REGION Network 21: Transition for STATE Num:60 StWtL1S2DownOver
   RUNG wire#powerrail
      Contact( #sStWtL1S2DownOver )
      I_Contact( #sStWtResetRel )
      Contact( #sSst )
      Contact( #iL1S2DownOver )
      Coil( #sStWtL1S2DownOver_T1 )
   END_RUNG
   // the same network as SCL:
   #sStWtL1S2DownOver_T1 := #sStWtL1S2DownOver AND NOT #sStWtResetRel AND #sSst AND #iL1S2DownOver;
END_REGION

REGION Network 22: STATE Num:60 StWtL1S2DownOver
   RUNG wire#powerrail
      Contact( #sStWtL1S2DownOver )
      wire#w1
      I_Contact( #sStWtResetRel )
      I_Contact( #sStWtL1S2DownOver_T1 )
      wire#w2
      Coil( #sStWtL1S2DownOver )
   END_RUNG
   RUNG wire#powerrail
      Contact( #sStWtLifterAtPos1_T1 )
   END_RUNG wire#w1
   RUNG wire#powerrail
      Contact( #sStRecovery_T7 )
   END_RUNG wire#w1
   RUNG wire#w2
      { S7_GenerateENO := "TRUE" } Move(in := 60, out1 => #StateNo)
   END_RUNG
   // the same network as SCL:
   #sStWtL1S2DownOver := (#sStWtL1S2DownOver OR #sStWtLifterAtPos1_T1 OR #sStRecovery_T7) AND NOT #sStWtResetRel AND NOT #sStWtL1S2DownOver_T1;
   IF #sStWtL1S2DownOver THEN #StateNo := 60; END_IF;
END_REGION

REGION Network 23: Actions for STATE Num:60 StWtL1S2DownOver
   RUNG wire#powerrail
      Contact( #sStWtL1S2DownOver )
      Coil( #qL1S2Down )
   END_RUNG
   // the same network as SCL:
   #qL1S2Down := #sStWtL1S2DownOver;
END_REGION

REGION Network 24: Transition for STATE Num:70 StWtOTSFrmConv
   RUNG wire#powerrail
      Contact( #sStWtOTSFrmConv )
      I_Contact( #sStWtResetRel )
      Contact( #sSst )
      Contact( #iOTSFrmConv )
      Coil( #sStWtOTSFrmConv_T1 )
   END_RUNG
   // the same network as SCL:
   #sStWtOTSFrmConv_T1 := #sStWtOTSFrmConv AND NOT #sStWtResetRel AND #sSst AND #iOTSFrmConv;
END_REGION

REGION Network 25: STATE Num:70 StWtOTSFrmConv
   RUNG wire#powerrail
      Contact( #sStWtOTSFrmConv )
      wire#w1
      I_Contact( #sStWtResetRel )
      I_Contact( #sStWtOTSFrmConv_T1 )
      wire#w2
      Coil( #sStWtOTSFrmConv )
   END_RUNG
   RUNG wire#powerrail
      Contact( #sStWtL1S2DownOver_T1 )
   END_RUNG wire#w1
   RUNG wire#w2
      { S7_GenerateENO := "TRUE" } Move(in := 70, out1 => #StateNo)
   END_RUNG
   // the same network as SCL:
   #sStWtOTSFrmConv := (#sStWtOTSFrmConv OR #sStWtL1S2DownOver_T1) AND NOT #sStWtResetRel AND NOT #sStWtOTSFrmConv_T1;
   IF #sStWtOTSFrmConv THEN #StateNo := 70; END_IF;
END_REGION

REGION Network 26: Actions for STATE Num:70 StWtOTSFrmConv
   RUNG wire#powerrail
      Contact( #sStWtOTSFrmConv )
      Coil( #qRTRToConv )
   END_RUNG
   // the same network as SCL:
   #qRTRToConv := #sStWtOTSFrmConv;
END_REGION

REGION Network 27: Transition for STATE Num:80 StWtL1RecvBegin
   RUNG wire#powerrail
      Contact( #sStWtL1RecvBegin )
      I_Contact( #sStWtResetRel )
      Contact( #sSst )
      I_Contact( #iReceiveAreaClear )
      Coil( #sStWtL1RecvBegin_T1 )
   END_RUNG
   // the same network as SCL:
   #sStWtL1RecvBegin_T1 := #sStWtL1RecvBegin AND NOT #sStWtResetRel AND #sSst AND NOT #iReceiveAreaClear;
END_REGION

REGION Network 28: STATE Num:80 StWtL1RecvBegin
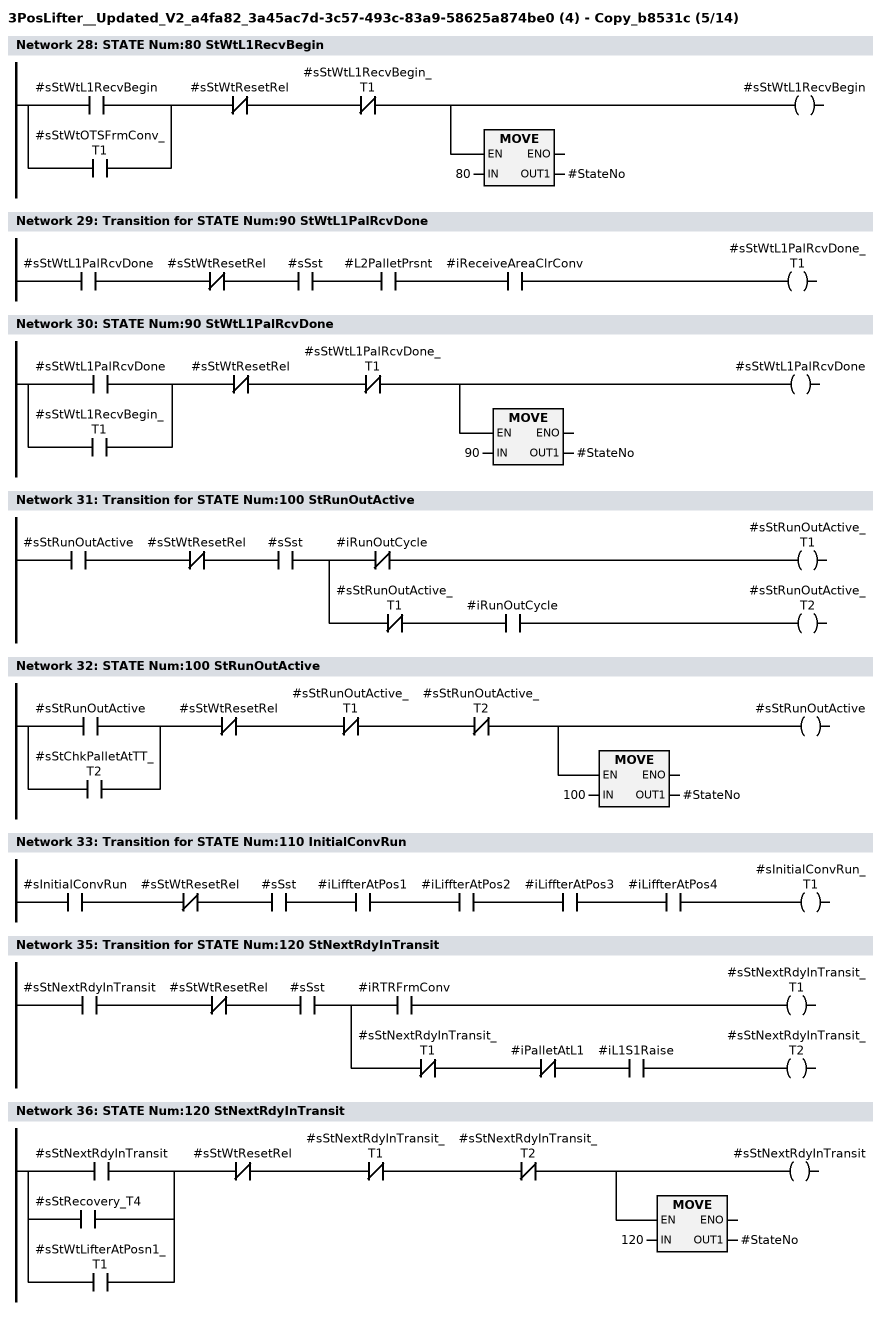
   RUNG wire#powerrail
      Contact( #sStWtL1RecvBegin )
      wire#w1
      I_Contact( #sStWtResetRel )
      I_Contact( #sStWtL1RecvBegin_T1 )
      wire#w2
      Coil( #sStWtL1RecvBegin )
   END_RUNG
   RUNG wire#powerrail
      Contact( #sStWtOTSFrmConv_T1 )
   END_RUNG wire#w1
   RUNG wire#w2
      { S7_GenerateENO := "TRUE" } Move(in := 80, out1 => #StateNo)
   END_RUNG
   // the same network as SCL:
   #sStWtL1RecvBegin := (#sStWtL1RecvBegin OR #sStWtOTSFrmConv_T1) AND NOT #sStWtResetRel AND NOT #sStWtL1RecvBegin_T1;
   IF #sStWtL1RecvBegin THEN #StateNo := 80; END_IF;
END_REGION

REGION Network 29: Transition for STATE Num:90 StWtL1PalRcvDone
   RUNG wire#powerrail
      Contact( #sStWtL1PalRcvDone )
      I_Contact( #sStWtResetRel )
      Contact( #sSst )
      Contact( #L2PalletPrsnt )
      Contact( #iReceiveAreaClrConv )
      Coil( #sStWtL1PalRcvDone_T1 )
   END_RUNG
   // the same network as SCL:
   #sStWtL1PalRcvDone_T1 := #sStWtL1PalRcvDone AND NOT #sStWtResetRel AND #sSst AND #L2PalletPrsnt AND #iReceiveAreaClrConv;
END_REGION

REGION Network 30: STATE Num:90 StWtL1PalRcvDone
   RUNG wire#powerrail
      Contact( #sStWtL1PalRcvDone )
      wire#w1
      I_Contact( #sStWtResetRel )
      I_Contact( #sStWtL1PalRcvDone_T1 )
      wire#w2
      Coil( #sStWtL1PalRcvDone )
   END_RUNG
   RUNG wire#powerrail
      Contact( #sStWtL1RecvBegin_T1 )
   END_RUNG wire#w1
   RUNG wire#w2
      { S7_GenerateENO := "TRUE" } Move(in := 90, out1 => #StateNo)
   END_RUNG
   // the same network as SCL:
   #sStWtL1PalRcvDone := (#sStWtL1PalRcvDone OR #sStWtL1RecvBegin_T1) AND NOT #sStWtResetRel AND NOT #sStWtL1PalRcvDone_T1;
   IF #sStWtL1PalRcvDone THEN #StateNo := 90; END_IF;
END_REGION

REGION Network 31: Transition for STATE Num:100 StRunOutActive
   RUNG wire#powerrail
      Contact( #sStRunOutActive )
      I_Contact( #sStWtResetRel )
      Contact( #sSst )
      wire#w1
      I_Contact( #iRunOutCycle )
      Coil( #sStRunOutActive_T1 )
   END_RUNG
   RUNG wire#w1
      I_Contact( #sStRunOutActive_T1 )
      Contact( #iRunOutCycle )
      Coil( #sStRunOutActive_T2 )
   END_RUNG
   // the same network as SCL:
   #_w1 := #sStRunOutActive AND NOT #sStWtResetRel AND #sSst;
   #sStRunOutActive_T1 := #_w1 AND NOT #iRunOutCycle;
   #sStRunOutActive_T2 := #_w1 AND NOT #sStRunOutActive_T1 AND #iRunOutCycle;
END_REGION

REGION Network 32: STATE Num:100 StRunOutActive
   RUNG wire#powerrail
      Contact( #sStRunOutActive )
      wire#w1
      I_Contact( #sStWtResetRel )
      I_Contact( #sStRunOutActive_T1 )
      I_Contact( #sStRunOutActive_T2 )
      wire#w2
      Coil( #sStRunOutActive )
   END_RUNG
   RUNG wire#powerrail
      Contact( #sStChkPalletAtTT_T2 )
   END_RUNG wire#w1
   RUNG wire#w2
      { S7_GenerateENO := "TRUE" } Move(in := 100, out1 => #StateNo)
   END_RUNG
   // the same network as SCL:
   #sStRunOutActive := (#sStRunOutActive OR #sStChkPalletAtTT_T2) AND NOT #sStWtResetRel AND NOT #sStRunOutActive_T1 AND NOT #sStRunOutActive_T2;
   IF #sStRunOutActive THEN #StateNo := 100; END_IF;
END_REGION

REGION Network 33: Transition for STATE Num:110 InitialConvRun
   RUNG wire#powerrail
      Contact( #sInitialConvRun )
      I_Contact( #sStWtResetRel )
      Contact( #sSst )
      Contact( #iLiffterAtPos1 )
      Contact( #iLiffterAtPos2 )
      Contact( #iLiffterAtPos3 )
      Contact( #iLiffterAtPos4 )
      Coil( #sInitialConvRun_T1 )
   END_RUNG
   // the same network as SCL:
   #sInitialConvRun_T1 := #sInitialConvRun AND NOT #sStWtResetRel AND #sSst AND #iLiffterAtPos1 AND #iLiffterAtPos2 AND #iLiffterAtPos3 AND #iLiffterAtPos4;
END_REGION

NETWORK
TITLE = STATE Num:110 InitialConvRun
      A(;
      O     #sInitialConvRun;
//wrong transition variable removed
      );
      AN    #sStWtResetRel;
      AN    #sInitialConvRun_T1;
      =     %L1.0;
      A     %L1.0;
      BLD   102;
      =     #sInitialConvRun;
      A     %L1.0;
      JNB   Label_110;
      L     110;
      T     #StateNo;
Label_110:NOP   0;

REGION Network 35: Transition for STATE Num:120 StNextRdyInTransit
   RUNG wire#powerrail
      Contact( #sStNextRdyInTransit )
      I_Contact( #sStWtResetRel )
      Contact( #sSst )
      wire#w1
      Contact( #iRTRFrmConv )
      Coil( #sStNextRdyInTransit_T1 )
   END_RUNG
   RUNG wire#w1
      I_Contact( #sStNextRdyInTransit_T1 )
      I_Contact( #iPalletAtL1 )
      Contact( #iL1S1Raise )
      Coil( #sStNextRdyInTransit_T2 )
   END_RUNG
   // the same network as SCL:
   #_w1 := #sStNextRdyInTransit AND NOT #sStWtResetRel AND #sSst;
   #sStNextRdyInTransit_T1 := #_w1 AND #iRTRFrmConv;
   #sStNextRdyInTransit_T2 := #_w1 AND NOT #sStNextRdyInTransit_T1 AND NOT #iPalletAtL1 AND #iL1S1Raise;
END_REGION

REGION Network 36: STATE Num:120 StNextRdyInTransit
   RUNG wire#powerrail
      Contact( #sStNextRdyInTransit )
      wire#w1
      I_Contact( #sStWtResetRel )
      I_Contact( #sStNextRdyInTransit_T1 )
      I_Contact( #sStNextRdyInTransit_T2 )
      wire#w2
      Coil( #sStNextRdyInTransit )
   END_RUNG
   RUNG wire#powerrail
      Contact( #sStRecovery_T4 )
   END_RUNG wire#w1
   RUNG wire#powerrail
      Contact( #sStWtLifterAtPosn1_T1 )
   END_RUNG wire#w1
   RUNG wire#w2
      { S7_GenerateENO := "TRUE" } Move(in := 120, out1 => #StateNo)
   END_RUNG
   // the same network as SCL:
   #sStNextRdyInTransit := (#sStNextRdyInTransit OR #sStRecovery_T4 OR #sStWtLifterAtPosn1_T1) AND NOT #sStWtResetRel AND NOT #sStNextRdyInTransit_T1 AND NOT #sStNextRdyInTransit_T2;
   IF #sStNextRdyInTransit THEN #StateNo := 120; END_IF;
END_REGION

REGION Network 37: Transition for STATE Num:130 StNextRdyInTransit_1
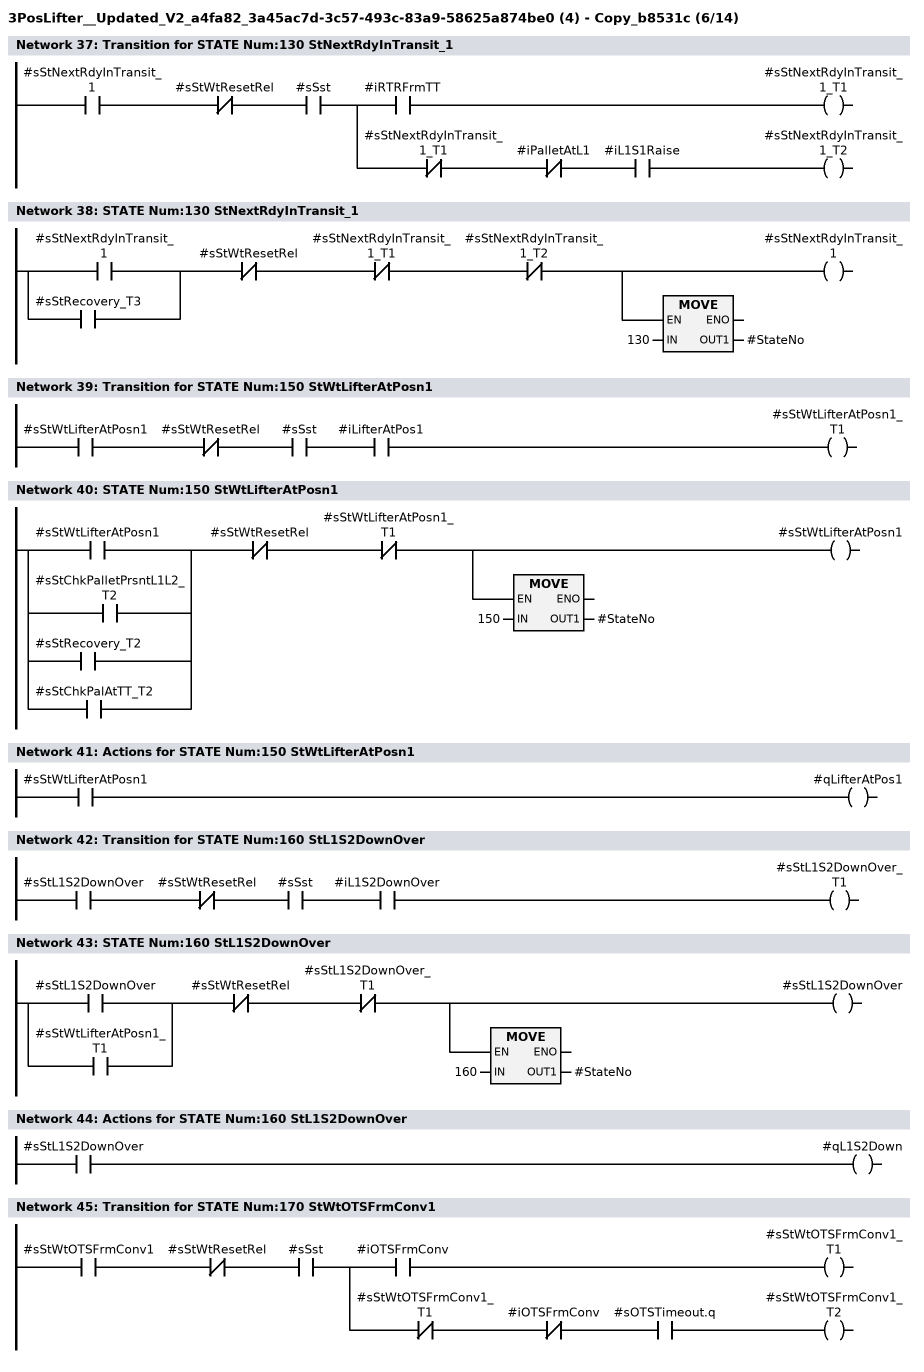
   RUNG wire#powerrail
      Contact( #sStNextRdyInTransit_1 )
      I_Contact( #sStWtResetRel )
      Contact( #sSst )
      wire#w1
      Contact( #iRTRFrmTT )
      Coil( #sStNextRdyInTransit_1_T1 )
   END_RUNG
   RUNG wire#w1
      I_Contact( #sStNextRdyInTransit_1_T1 )
      I_Contact( #iPalletAtL1 )
      Contact( #iL1S1Raise )
      Coil( #sStNextRdyInTransit_1_T2 )
   END_RUNG
   // the same network as SCL:
   #_w1 := #sStNextRdyInTransit_1 AND NOT #sStWtResetRel AND #sSst;
   #sStNextRdyInTransit_1_T1 := #_w1 AND #iRTRFrmTT;
   #sStNextRdyInTransit_1_T2 := #_w1 AND NOT #sStNextRdyInTransit_1_T1 AND NOT #iPalletAtL1 AND #iL1S1Raise;
END_REGION

REGION Network 38: STATE Num:130 StNextRdyInTransit_1
   RUNG wire#powerrail
      Contact( #sStNextRdyInTransit_1 )
      wire#w1
      I_Contact( #sStWtResetRel )
      I_Contact( #sStNextRdyInTransit_1_T1 )
      I_Contact( #sStNextRdyInTransit_1_T2 )
      wire#w2
      Coil( #sStNextRdyInTransit_1 )
   END_RUNG
   RUNG wire#powerrail
      Contact( #sStRecovery_T3 )
   END_RUNG wire#w1
   RUNG wire#w2
      { S7_GenerateENO := "TRUE" } Move(in := 130, out1 => #StateNo)
   END_RUNG
   // the same network as SCL:
   #sStNextRdyInTransit_1 := (#sStNextRdyInTransit_1 OR #sStRecovery_T3) AND NOT #sStWtResetRel AND NOT #sStNextRdyInTransit_1_T1 AND NOT #sStNextRdyInTransit_1_T2;
   IF #sStNextRdyInTransit_1 THEN #StateNo := 130; END_IF;
END_REGION

REGION Network 39: Transition for STATE Num:150 StWtLifterAtPosn1
   RUNG wire#powerrail
      Contact( #sStWtLifterAtPosn1 )
      I_Contact( #sStWtResetRel )
      Contact( #sSst )
      Contact( #iLifterAtPos1 )
      Coil( #sStWtLifterAtPosn1_T1 )
   END_RUNG
   // the same network as SCL:
   #sStWtLifterAtPosn1_T1 := #sStWtLifterAtPosn1 AND NOT #sStWtResetRel AND #sSst AND #iLifterAtPos1;
END_REGION

REGION Network 40: STATE Num:150 StWtLifterAtPosn1
   RUNG wire#powerrail
      Contact( #sStWtLifterAtPosn1 )
      wire#w1
      I_Contact( #sStWtResetRel )
      I_Contact( #sStWtLifterAtPosn1_T1 )
      wire#w2
      Coil( #sStWtLifterAtPosn1 )
   END_RUNG
   RUNG wire#powerrail
      Contact( #sStChkPalletPrsntL1L2_T2 )
   END_RUNG wire#w1
   RUNG wire#powerrail
      Contact( #sStRecovery_T2 )
   END_RUNG wire#w1
   RUNG wire#powerrail
      Contact( #sStChkPalAtTT_T2 )
   END_RUNG wire#w1
   RUNG wire#w2
      { S7_GenerateENO := "TRUE" } Move(in := 150, out1 => #StateNo)
   END_RUNG
   // the same network as SCL:
   #sStWtLifterAtPosn1 := (#sStWtLifterAtPosn1 OR #sStChkPalletPrsntL1L2_T2 OR #sStRecovery_T2 OR #sStChkPalAtTT_T2) AND NOT #sStWtResetRel AND NOT #sStWtLifterAtPosn1_T1;
   IF #sStWtLifterAtPosn1 THEN #StateNo := 150; END_IF;
END_REGION

REGION Network 41: Actions for STATE Num:150 StWtLifterAtPosn1
   RUNG wire#powerrail
      Contact( #sStWtLifterAtPosn1 )
      Coil( #qLifterAtPos1 )
   END_RUNG
   // the same network as SCL:
   #qLifterAtPos1 := #sStWtLifterAtPosn1;
END_REGION

REGION Network 42: Transition for STATE Num:160 StL1S2DownOver
   RUNG wire#powerrail
      Contact( #sStL1S2DownOver )
      I_Contact( #sStWtResetRel )
      Contact( #sSst )
      Contact( #iL1S2DownOver )
      Coil( #sStL1S2DownOver_T1 )
   END_RUNG
   // the same network as SCL:
   #sStL1S2DownOver_T1 := #sStL1S2DownOver AND NOT #sStWtResetRel AND #sSst AND #iL1S2DownOver;
END_REGION

REGION Network 43: STATE Num:160 StL1S2DownOver
   RUNG wire#powerrail
      Contact( #sStL1S2DownOver )
      wire#w1
      I_Contact( #sStWtResetRel )
      I_Contact( #sStL1S2DownOver_T1 )
      wire#w2
      Coil( #sStL1S2DownOver )
   END_RUNG
   RUNG wire#powerrail
      Contact( #sStWtLifterAtPosn1_T1 )
   END_RUNG wire#w1
   RUNG wire#w2
      { S7_GenerateENO := "TRUE" } Move(in := 160, out1 => #StateNo)
   END_RUNG
   // the same network as SCL:
   #sStL1S2DownOver := (#sStL1S2DownOver OR #sStWtLifterAtPosn1_T1) AND NOT #sStWtResetRel AND NOT #sStL1S2DownOver_T1;
   IF #sStL1S2DownOver THEN #StateNo := 160; END_IF;
END_REGION

REGION Network 44: Actions for STATE Num:160 StL1S2DownOver
   RUNG wire#powerrail
      Contact( #sStL1S2DownOver )
      Coil( #qL1S2Down )
   END_RUNG
   // the same network as SCL:
   #qL1S2Down := #sStL1S2DownOver;
END_REGION

REGION Network 45: Transition for STATE Num:170 StWtOTSFrmConv1
   RUNG wire#powerrail
      Contact( #sStWtOTSFrmConv1 )
      I_Contact( #sStWtResetRel )
      Contact( #sSst )
      wire#w1
      Contact( #iOTSFrmConv )
      Coil( #sStWtOTSFrmConv1_T1 )
   END_RUNG
   RUNG wire#w1
      I_Contact( #sStWtOTSFrmConv1_T1 )
      I_Contact( #iOTSFrmConv )
      Contact( #sOTSTimeout.q )
      Coil( #sStWtOTSFrmConv1_T2 )
   END_RUNG
   // the same network as SCL:
   #_w1 := #sStWtOTSFrmConv1 AND NOT #sStWtResetRel AND #sSst;
   #sStWtOTSFrmConv1_T1 := #_w1 AND #iOTSFrmConv;
   #sStWtOTSFrmConv1_T2 := #_w1 AND NOT #sStWtOTSFrmConv1_T1 AND NOT #iOTSFrmConv AND #sOTSTimeout.q;
END_REGION

REGION Network 46: STATE Num:170 StWtOTSFrmConv1
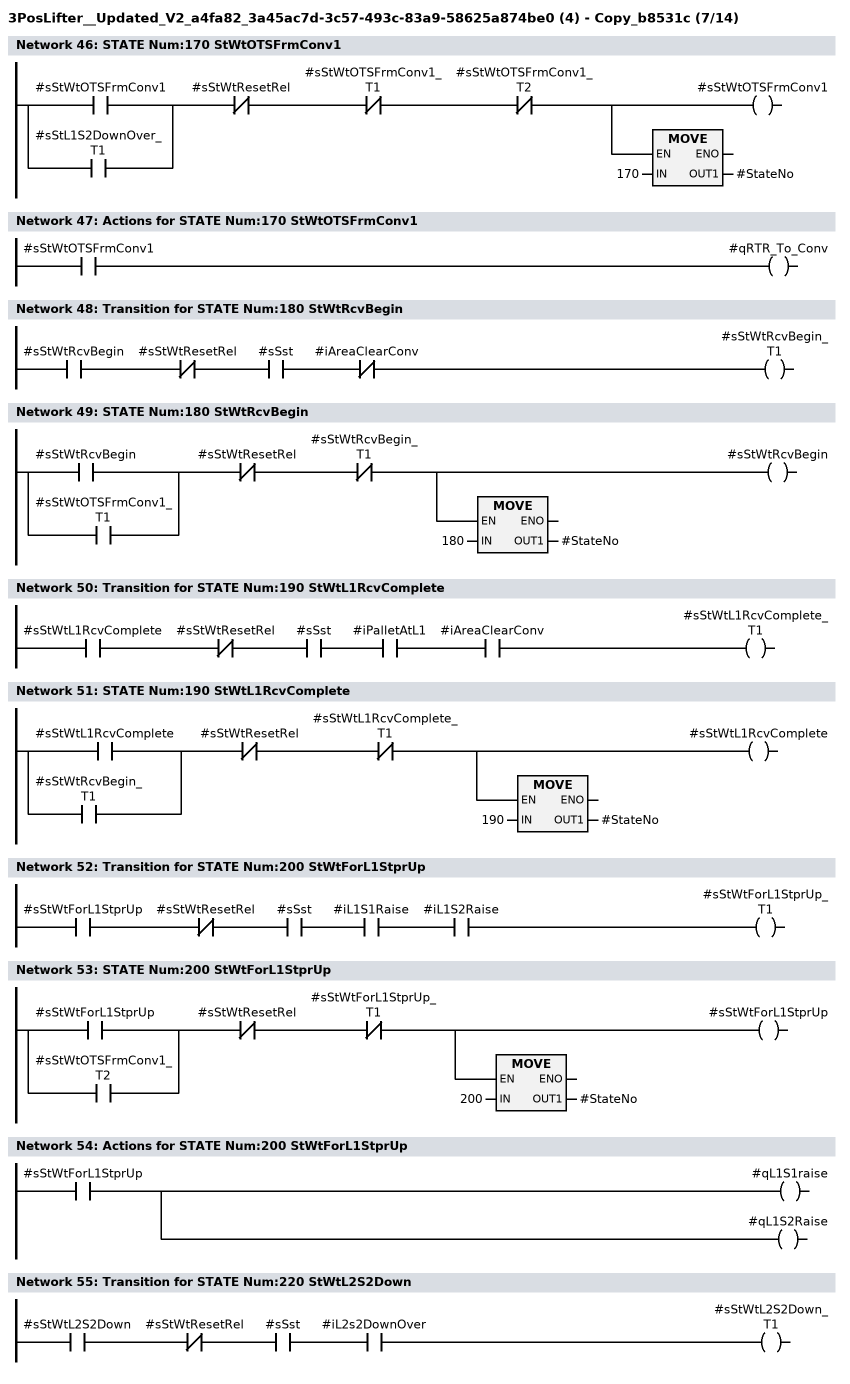
   RUNG wire#powerrail
      Contact( #sStWtOTSFrmConv1 )
      wire#w1
      I_Contact( #sStWtResetRel )
      I_Contact( #sStWtOTSFrmConv1_T1 )
      I_Contact( #sStWtOTSFrmConv1_T2 )
      wire#w2
      Coil( #sStWtOTSFrmConv1 )
   END_RUNG
   RUNG wire#powerrail
      Contact( #sStL1S2DownOver_T1 )
   END_RUNG wire#w1
   RUNG wire#w2
      { S7_GenerateENO := "TRUE" } Move(in := 170, out1 => #StateNo)
   END_RUNG
   // the same network as SCL:
   #sStWtOTSFrmConv1 := (#sStWtOTSFrmConv1 OR #sStL1S2DownOver_T1) AND NOT #sStWtResetRel AND NOT #sStWtOTSFrmConv1_T1 AND NOT #sStWtOTSFrmConv1_T2;
   IF #sStWtOTSFrmConv1 THEN #StateNo := 170; END_IF;
END_REGION

REGION Network 47: Actions for STATE Num:170 StWtOTSFrmConv1
   RUNG wire#powerrail
      Contact( #sStWtOTSFrmConv1 )
      Coil( #qRTR_To_Conv )
   END_RUNG
   // the same network as SCL:
   #qRTR_To_Conv := #sStWtOTSFrmConv1;
END_REGION

REGION Network 48: Transition for STATE Num:180 StWtRcvBegin
   RUNG wire#powerrail
      Contact( #sStWtRcvBegin )
      I_Contact( #sStWtResetRel )
      Contact( #sSst )
      I_Contact( #iAreaClearConv )
      Coil( #sStWtRcvBegin_T1 )
   END_RUNG
   // the same network as SCL:
   #sStWtRcvBegin_T1 := #sStWtRcvBegin AND NOT #sStWtResetRel AND #sSst AND NOT #iAreaClearConv;
END_REGION

REGION Network 49: STATE Num:180 StWtRcvBegin
   RUNG wire#powerrail
      Contact( #sStWtRcvBegin )
      wire#w1
      I_Contact( #sStWtResetRel )
      I_Contact( #sStWtRcvBegin_T1 )
      wire#w2
      Coil( #sStWtRcvBegin )
   END_RUNG
   RUNG wire#powerrail
      Contact( #sStWtOTSFrmConv1_T1 )
   END_RUNG wire#w1
   RUNG wire#w2
      { S7_GenerateENO := "TRUE" } Move(in := 180, out1 => #StateNo)
   END_RUNG
   // the same network as SCL:
   #sStWtRcvBegin := (#sStWtRcvBegin OR #sStWtOTSFrmConv1_T1) AND NOT #sStWtResetRel AND NOT #sStWtRcvBegin_T1;
   IF #sStWtRcvBegin THEN #StateNo := 180; END_IF;
END_REGION

REGION Network 50: Transition for STATE Num:190 StWtL1RcvComplete
   RUNG wire#powerrail
      Contact( #sStWtL1RcvComplete )
      I_Contact( #sStWtResetRel )
      Contact( #sSst )
      Contact( #iPalletAtL1 )
      Contact( #iAreaClearConv )
      Coil( #sStWtL1RcvComplete_T1 )
   END_RUNG
   // the same network as SCL:
   #sStWtL1RcvComplete_T1 := #sStWtL1RcvComplete AND NOT #sStWtResetRel AND #sSst AND #iPalletAtL1 AND #iAreaClearConv;
END_REGION

REGION Network 51: STATE Num:190 StWtL1RcvComplete
   RUNG wire#powerrail
      Contact( #sStWtL1RcvComplete )
      wire#w1
      I_Contact( #sStWtResetRel )
      I_Contact( #sStWtL1RcvComplete_T1 )
      wire#w2
      Coil( #sStWtL1RcvComplete )
   END_RUNG
   RUNG wire#powerrail
      Contact( #sStWtRcvBegin_T1 )
   END_RUNG wire#w1
   RUNG wire#w2
      { S7_GenerateENO := "TRUE" } Move(in := 190, out1 => #StateNo)
   END_RUNG
   // the same network as SCL:
   #sStWtL1RcvComplete := (#sStWtL1RcvComplete OR #sStWtRcvBegin_T1) AND NOT #sStWtResetRel AND NOT #sStWtL1RcvComplete_T1;
   IF #sStWtL1RcvComplete THEN #StateNo := 190; END_IF;
END_REGION

REGION Network 52: Transition for STATE Num:200 StWtForL1StprUp
   RUNG wire#powerrail
      Contact( #sStWtForL1StprUp )
      I_Contact( #sStWtResetRel )
      Contact( #sSst )
      Contact( #iL1S1Raise )
      Contact( #iL1S2Raise )
      Coil( #sStWtForL1StprUp_T1 )
   END_RUNG
   // the same network as SCL:
   #sStWtForL1StprUp_T1 := #sStWtForL1StprUp AND NOT #sStWtResetRel AND #sSst AND #iL1S1Raise AND #iL1S2Raise;
END_REGION

REGION Network 53: STATE Num:200 StWtForL1StprUp
   RUNG wire#powerrail
      Contact( #sStWtForL1StprUp )
      wire#w1
      I_Contact( #sStWtResetRel )
      I_Contact( #sStWtForL1StprUp_T1 )
      wire#w2
      Coil( #sStWtForL1StprUp )
   END_RUNG
   RUNG wire#powerrail
      Contact( #sStWtOTSFrmConv1_T2 )
   END_RUNG wire#w1
   RUNG wire#w2
      { S7_GenerateENO := "TRUE" } Move(in := 200, out1 => #StateNo)
   END_RUNG
   // the same network as SCL:
   #sStWtForL1StprUp := (#sStWtForL1StprUp OR #sStWtOTSFrmConv1_T2) AND NOT #sStWtResetRel AND NOT #sStWtForL1StprUp_T1;
   IF #sStWtForL1StprUp THEN #StateNo := 200; END_IF;
END_REGION

REGION Network 54: Actions for STATE Num:200 StWtForL1StprUp
   RUNG wire#powerrail
      Contact( #sStWtForL1StprUp )
      wire#w1
      Coil( #qL1S1raise )
   END_RUNG
   RUNG wire#w1
      Coil( #qL1S2Raise )
   END_RUNG
   // the same network as SCL:
   #qL1S1raise := #sStWtForL1StprUp;
   #qL1S2Raise := #sStWtForL1StprUp;
END_REGION

REGION Network 55: Transition for STATE Num:220 StWtL2S2Down
   RUNG wire#powerrail
      Contact( #sStWtL2S2Down )
      I_Contact( #sStWtResetRel )
      Contact( #sSst )
      Contact( #iL2s2DownOver )
      Coil( #sStWtL2S2Down_T1 )
   END_RUNG
   // the same network as SCL:
   #sStWtL2S2Down_T1 := #sStWtL2S2Down AND NOT #sStWtResetRel AND #sSst AND #iL2s2DownOver;
END_REGION

REGION Network 56: STATE Num:220 StWtL2S2Down
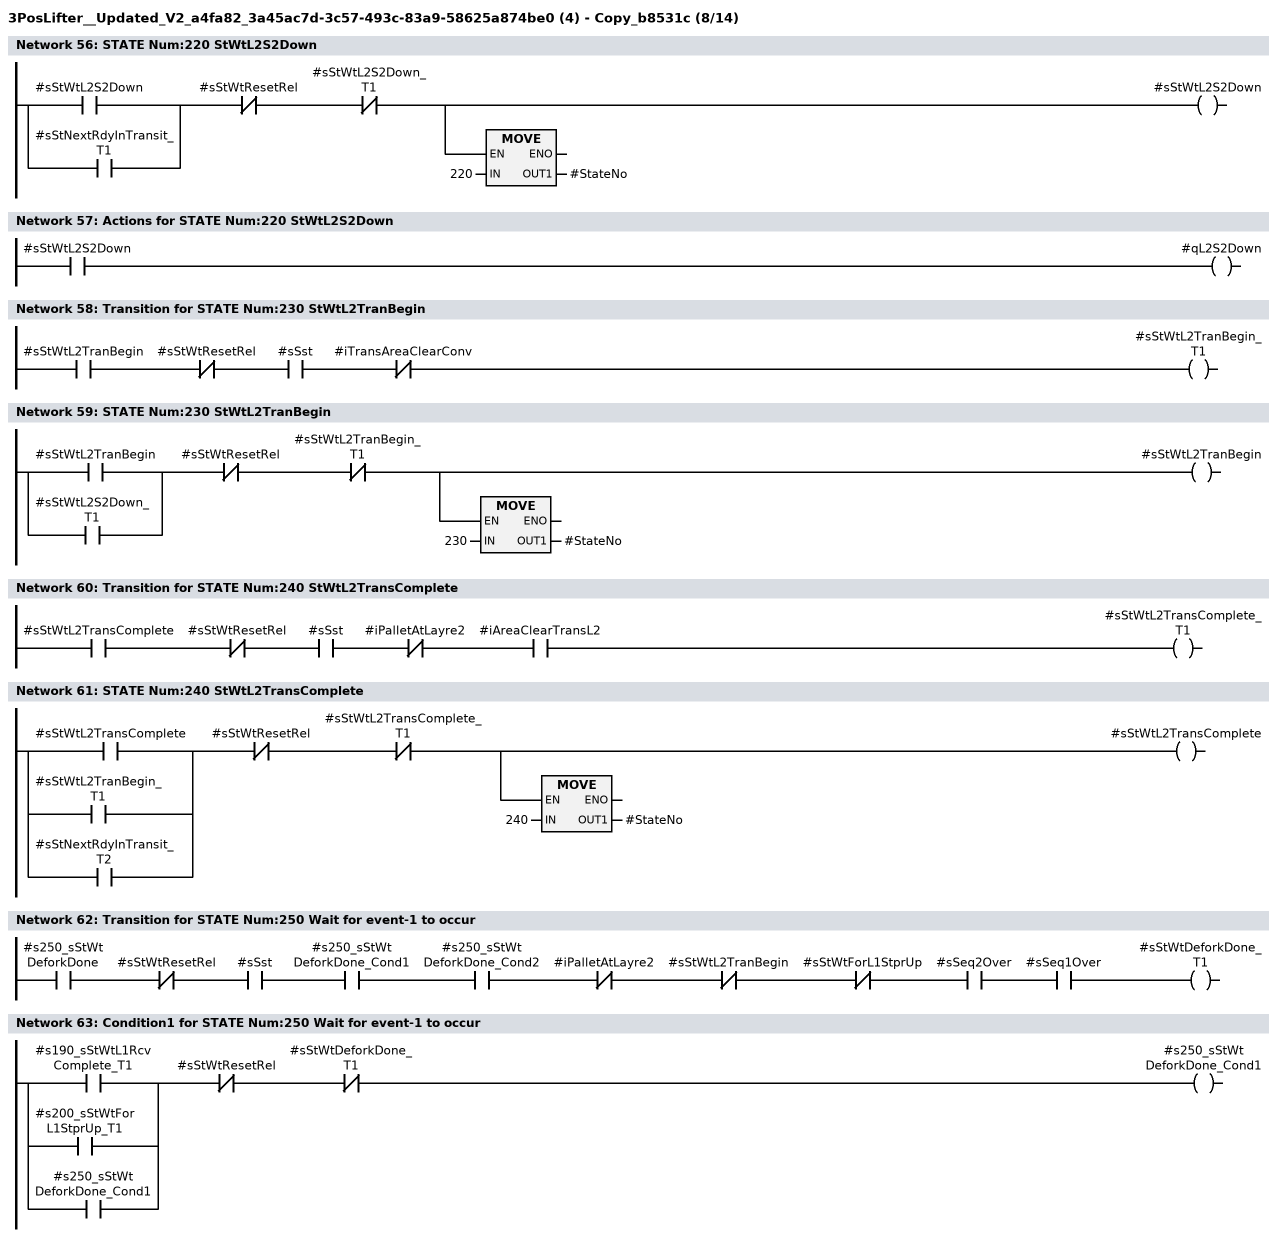
   RUNG wire#powerrail
      Contact( #sStWtL2S2Down )
      wire#w1
      I_Contact( #sStWtResetRel )
      I_Contact( #sStWtL2S2Down_T1 )
      wire#w2
      Coil( #sStWtL2S2Down )
   END_RUNG
   RUNG wire#powerrail
      Contact( #sStNextRdyInTransit_T1 )
   END_RUNG wire#w1
   RUNG wire#w2
      { S7_GenerateENO := "TRUE" } Move(in := 220, out1 => #StateNo)
   END_RUNG
   // the same network as SCL:
   #sStWtL2S2Down := (#sStWtL2S2Down OR #sStNextRdyInTransit_T1) AND NOT #sStWtResetRel AND NOT #sStWtL2S2Down_T1;
   IF #sStWtL2S2Down THEN #StateNo := 220; END_IF;
END_REGION

REGION Network 57: Actions for STATE Num:220 StWtL2S2Down
   RUNG wire#powerrail
      Contact( #sStWtL2S2Down )
      Coil( #qL2S2Down )
   END_RUNG
   // the same network as SCL:
   #qL2S2Down := #sStWtL2S2Down;
END_REGION

REGION Network 58: Transition for STATE Num:230 StWtL2TranBegin
   RUNG wire#powerrail
      Contact( #sStWtL2TranBegin )
      I_Contact( #sStWtResetRel )
      Contact( #sSst )
      I_Contact( #iTransAreaClearConv )
      Coil( #sStWtL2TranBegin_T1 )
   END_RUNG
   // the same network as SCL:
   #sStWtL2TranBegin_T1 := #sStWtL2TranBegin AND NOT #sStWtResetRel AND #sSst AND NOT #iTransAreaClearConv;
END_REGION

REGION Network 59: STATE Num:230 StWtL2TranBegin
   RUNG wire#powerrail
      Contact( #sStWtL2TranBegin )
      wire#w1
      I_Contact( #sStWtResetRel )
      I_Contact( #sStWtL2TranBegin_T1 )
      wire#w2
      Coil( #sStWtL2TranBegin )
   END_RUNG
   RUNG wire#powerrail
      Contact( #sStWtL2S2Down_T1 )
   END_RUNG wire#w1
   RUNG wire#w2
      { S7_GenerateENO := "TRUE" } Move(in := 230, out1 => #StateNo)
   END_RUNG
   // the same network as SCL:
   #sStWtL2TranBegin := (#sStWtL2TranBegin OR #sStWtL2S2Down_T1) AND NOT #sStWtResetRel AND NOT #sStWtL2TranBegin_T1;
   IF #sStWtL2TranBegin THEN #StateNo := 230; END_IF;
END_REGION

REGION Network 60: Transition for STATE Num:240 StWtL2TransComplete
   RUNG wire#powerrail
      Contact( #sStWtL2TransComplete )
      I_Contact( #sStWtResetRel )
      Contact( #sSst )
      I_Contact( #iPalletAtLayre2 )
      Contact( #iAreaClearTransL2 )
      Coil( #sStWtL2TransComplete_T1 )
   END_RUNG
   // the same network as SCL:
   #sStWtL2TransComplete_T1 := #sStWtL2TransComplete AND NOT #sStWtResetRel AND #sSst AND NOT #iPalletAtLayre2 AND #iAreaClearTransL2;
END_REGION

REGION Network 61: STATE Num:240 StWtL2TransComplete
   RUNG wire#powerrail
      Contact( #sStWtL2TransComplete )
      wire#w1
      I_Contact( #sStWtResetRel )
      I_Contact( #sStWtL2TransComplete_T1 )
      wire#w2
      Coil( #sStWtL2TransComplete )
   END_RUNG
   RUNG wire#powerrail
      Contact( #sStWtL2TranBegin_T1 )
   END_RUNG wire#w1
   RUNG wire#powerrail
      Contact( #sStNextRdyInTransit_T2 )
   END_RUNG wire#w1
   RUNG wire#w2
      { S7_GenerateENO := "TRUE" } Move(in := 240, out1 => #StateNo)
   END_RUNG
   // the same network as SCL:
   #sStWtL2TransComplete := (#sStWtL2TransComplete OR #sStWtL2TranBegin_T1 OR #sStNextRdyInTransit_T2) AND NOT #sStWtResetRel AND NOT #sStWtL2TransComplete_T1;
   IF #sStWtL2TransComplete THEN #StateNo := 240; END_IF;
END_REGION

REGION Network 62: Transition for STATE Num:250 Wait for event-1 to occur
   RUNG wire#powerrail
      Contact( #s250_sStWtDeforkDone )
      I_Contact( #sStWtResetRel )
      Contact( #sSst )
      Contact( #s250_sStWtDeforkDone_Cond1 )
      Contact( #s250_sStWtDeforkDone_Cond2 )
      I_Contact( #iPalletAtLayre2 )
      I_Contact( #sStWtL2TranBegin )
      I_Contact( #sStWtForL1StprUp )
      Contact( #sSeq2Over )
      Contact( #sSeq1Over )
      Coil( #sStWtDeforkDone_T1 )
   END_RUNG
   // the same network as SCL:
   #sStWtDeforkDone_T1 := #s250_sStWtDeforkDone AND NOT #sStWtResetRel AND #sSst AND #s250_sStWtDeforkDone_Cond1 AND #s250_sStWtDeforkDone_Cond2 AND NOT #iPalletAtLayre2 AND NOT #sStWtL2TranBegin AND NOT #sStWtForL1StprUp AND #sSeq2Over AND #sSeq1Over;
END_REGION

REGION Network 63: Condition1 for STATE Num:250 Wait for event-1 to occur
   RUNG wire#powerrail
      Contact( #s190_sStWtL1RcvComplete_T1 )
      wire#w1
      I_Contact( #sStWtResetRel )
      I_Contact( #sStWtDeforkDone_T1 )
      Coil( #s250_sStWtDeforkDone_Cond1 )
   END_RUNG
   RUNG wire#powerrail
      Contact( #s200_sStWtForL1StprUp_T1 )
   END_RUNG wire#w1
   RUNG wire#powerrail
      Contact( #s250_sStWtDeforkDone_Cond1 )
   END_RUNG wire#w1
   // the same network as SCL:
   #s250_sStWtDeforkDone_Cond1 := (#s190_sStWtL1RcvComplete_T1 OR #s200_sStWtForL1StprUp_T1 OR #s250_sStWtDeforkDone_Cond1) AND NOT #sStWtResetRel AND NOT #sStWtDeforkDone_T1;
END_REGION

REGION Network 64: Condition2 for STATE Num:250 Wait for event-1 to occur
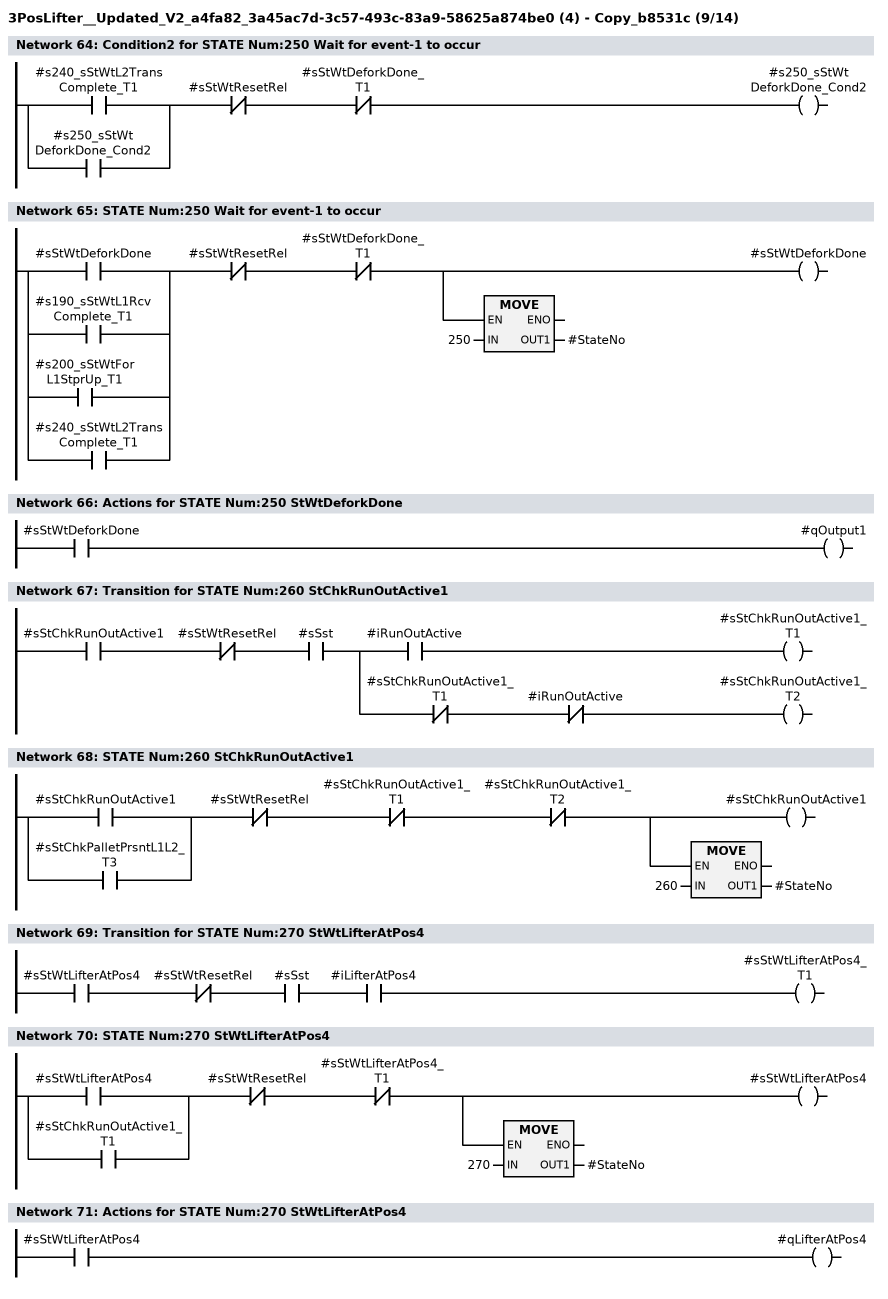
   RUNG wire#powerrail
      Contact( #s240_sStWtL2TransComplete_T1 )
      wire#w1
      I_Contact( #sStWtResetRel )
      I_Contact( #sStWtDeforkDone_T1 )
      Coil( #s250_sStWtDeforkDone_Cond2 )
   END_RUNG
   RUNG wire#powerrail
      Contact( #s250_sStWtDeforkDone_Cond2 )
   END_RUNG wire#w1
   // the same network as SCL:
   #s250_sStWtDeforkDone_Cond2 := (#s240_sStWtL2TransComplete_T1 OR #s250_sStWtDeforkDone_Cond2) AND NOT #sStWtResetRel AND NOT #sStWtDeforkDone_T1;
END_REGION

REGION Network 65: STATE Num:250 Wait for event-1 to occur
   RUNG wire#powerrail
      Contact( #sStWtDeforkDone )
      wire#w1
      I_Contact( #sStWtResetRel )
      I_Contact( #sStWtDeforkDone_T1 )
      wire#w2
      Coil( #sStWtDeforkDone )
   END_RUNG
   RUNG wire#powerrail
      Contact( #s190_sStWtL1RcvComplete_T1 )
   END_RUNG wire#w1
   RUNG wire#powerrail
      Contact( #s200_sStWtForL1StprUp_T1 )
   END_RUNG wire#w1
   RUNG wire#powerrail
      Contact( #s240_sStWtL2TransComplete_T1 )
   END_RUNG wire#w1
   RUNG wire#w2
      { S7_GenerateENO := "TRUE" } Move(in := 250, out1 => #StateNo)
   END_RUNG
   // the same network as SCL:
   #sStWtDeforkDone := (#sStWtDeforkDone OR #s190_sStWtL1RcvComplete_T1 OR #s200_sStWtForL1StprUp_T1 OR #s240_sStWtL2TransComplete_T1) AND NOT #sStWtResetRel AND NOT #sStWtDeforkDone_T1;
   IF #sStWtDeforkDone THEN #StateNo := 250; END_IF;
END_REGION

REGION Network 66: Actions for STATE Num:250 StWtDeforkDone
   RUNG wire#powerrail
      Contact( #sStWtDeforkDone )
      Coil( #qOutput1 )
   END_RUNG
   // the same network as SCL:
   #qOutput1 := #sStWtDeforkDone;
END_REGION

REGION Network 67: Transition for STATE Num:260 StChkRunOutActive1
   RUNG wire#powerrail
      Contact( #sStChkRunOutActive1 )
      I_Contact( #sStWtResetRel )
      Contact( #sSst )
      wire#w1
      Contact( #iRunOutActive )
      Coil( #sStChkRunOutActive1_T1 )
   END_RUNG
   RUNG wire#w1
      I_Contact( #sStChkRunOutActive1_T1 )
      I_Contact( #iRunOutActive )
      Coil( #sStChkRunOutActive1_T2 )
   END_RUNG
   // the same network as SCL:
   #_w1 := #sStChkRunOutActive1 AND NOT #sStWtResetRel AND #sSst;
   #sStChkRunOutActive1_T1 := #_w1 AND #iRunOutActive;
   #sStChkRunOutActive1_T2 := #_w1 AND NOT #sStChkRunOutActive1_T1 AND NOT #iRunOutActive;
END_REGION

REGION Network 68: STATE Num:260 StChkRunOutActive1
   RUNG wire#powerrail
      Contact( #sStChkRunOutActive1 )
      wire#w1
      I_Contact( #sStWtResetRel )
      I_Contact( #sStChkRunOutActive1_T1 )
      I_Contact( #sStChkRunOutActive1_T2 )
      wire#w2
      Coil( #sStChkRunOutActive1 )
   END_RUNG
   RUNG wire#powerrail
      Contact( #sStChkPalletPrsntL1L2_T3 )
   END_RUNG wire#w1
   RUNG wire#w2
      { S7_GenerateENO := "TRUE" } Move(in := 260, out1 => #StateNo)
   END_RUNG
   // the same network as SCL:
   #sStChkRunOutActive1 := (#sStChkRunOutActive1 OR #sStChkPalletPrsntL1L2_T3) AND NOT #sStWtResetRel AND NOT #sStChkRunOutActive1_T1 AND NOT #sStChkRunOutActive1_T2;
   IF #sStChkRunOutActive1 THEN #StateNo := 260; END_IF;
END_REGION

REGION Network 69: Transition for STATE Num:270 StWtLifterAtPos4
   RUNG wire#powerrail
      Contact( #sStWtLifterAtPos4 )
      I_Contact( #sStWtResetRel )
      Contact( #sSst )
      Contact( #iLifterAtPos4 )
      Coil( #sStWtLifterAtPos4_T1 )
   END_RUNG
   // the same network as SCL:
   #sStWtLifterAtPos4_T1 := #sStWtLifterAtPos4 AND NOT #sStWtResetRel AND #sSst AND #iLifterAtPos4;
END_REGION

REGION Network 70: STATE Num:270 StWtLifterAtPos4
   RUNG wire#powerrail
      Contact( #sStWtLifterAtPos4 )
      wire#w1
      I_Contact( #sStWtResetRel )
      I_Contact( #sStWtLifterAtPos4_T1 )
      wire#w2
      Coil( #sStWtLifterAtPos4 )
   END_RUNG
   RUNG wire#powerrail
      Contact( #sStChkRunOutActive1_T1 )
   END_RUNG wire#w1
   RUNG wire#w2
      { S7_GenerateENO := "TRUE" } Move(in := 270, out1 => #StateNo)
   END_RUNG
   // the same network as SCL:
   #sStWtLifterAtPos4 := (#sStWtLifterAtPos4 OR #sStChkRunOutActive1_T1) AND NOT #sStWtResetRel AND NOT #sStWtLifterAtPos4_T1;
   IF #sStWtLifterAtPos4 THEN #StateNo := 270; END_IF;
END_REGION

REGION Network 71: Actions for STATE Num:270 StWtLifterAtPos4
   RUNG wire#powerrail
      Contact( #sStWtLifterAtPos4 )
      Coil( #qLifterAtPos4 )
   END_RUNG
   // the same network as SCL:
   #qLifterAtPos4 := #sStWtLifterAtPos4;
END_REGION

REGION Network 72: Transition for STATE Num:280 StWtRTRFrmConvPos4
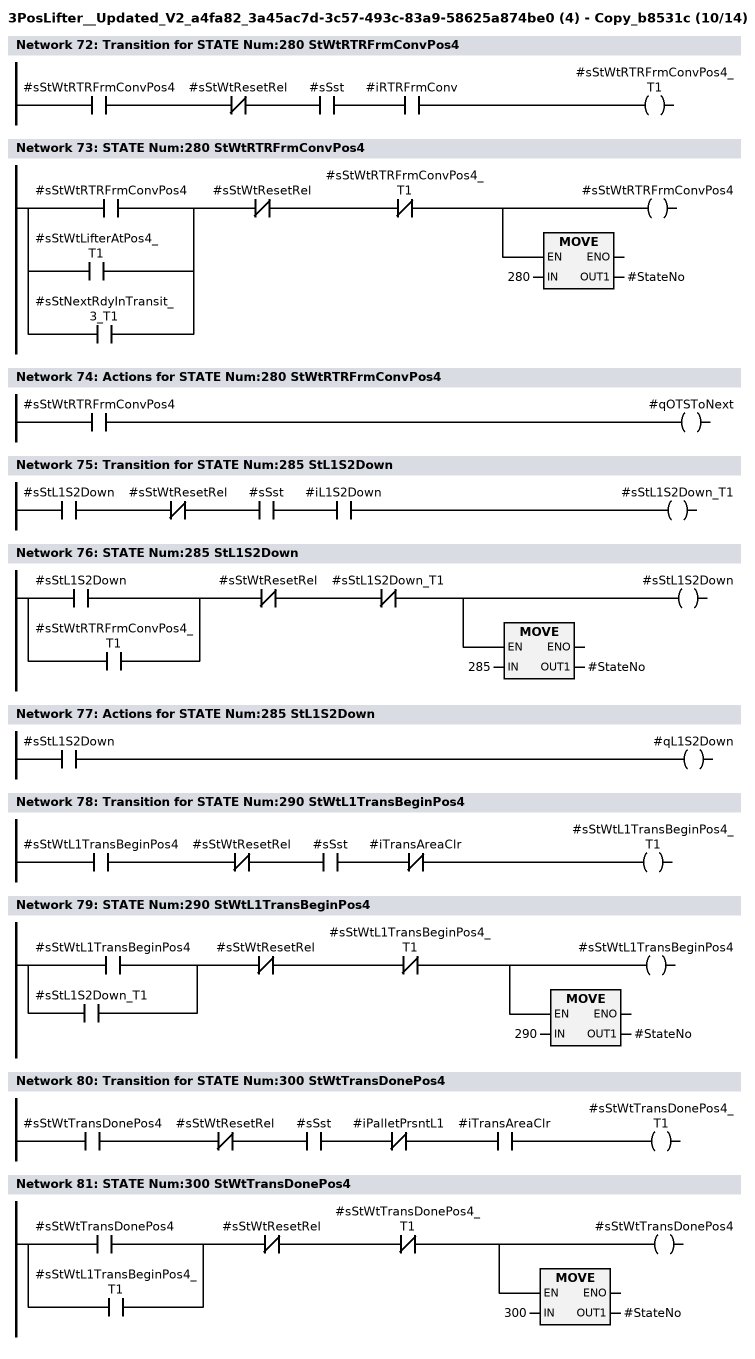
   RUNG wire#powerrail
      Contact( #sStWtRTRFrmConvPos4 )
      I_Contact( #sStWtResetRel )
      Contact( #sSst )
      Contact( #iRTRFrmConv )
      Coil( #sStWtRTRFrmConvPos4_T1 )
   END_RUNG
   // the same network as SCL:
   #sStWtRTRFrmConvPos4_T1 := #sStWtRTRFrmConvPos4 AND NOT #sStWtResetRel AND #sSst AND #iRTRFrmConv;
END_REGION

REGION Network 73: STATE Num:280 StWtRTRFrmConvPos4
   RUNG wire#powerrail
      Contact( #sStWtRTRFrmConvPos4 )
      wire#w1
      I_Contact( #sStWtResetRel )
      I_Contact( #sStWtRTRFrmConvPos4_T1 )
      wire#w2
      Coil( #sStWtRTRFrmConvPos4 )
   END_RUNG
   RUNG wire#powerrail
      Contact( #sStWtLifterAtPos4_T1 )
   END_RUNG wire#w1
   RUNG wire#powerrail
      Contact( #sStNextRdyInTransit_3_T1 )
   END_RUNG wire#w1
   RUNG wire#w2
      { S7_GenerateENO := "TRUE" } Move(in := 280, out1 => #StateNo)
   END_RUNG
   // the same network as SCL:
   #sStWtRTRFrmConvPos4 := (#sStWtRTRFrmConvPos4 OR #sStWtLifterAtPos4_T1 OR #sStNextRdyInTransit_3_T1) AND NOT #sStWtResetRel AND NOT #sStWtRTRFrmConvPos4_T1;
   IF #sStWtRTRFrmConvPos4 THEN #StateNo := 280; END_IF;
END_REGION

REGION Network 74: Actions for STATE Num:280 StWtRTRFrmConvPos4
   RUNG wire#powerrail
      Contact( #sStWtRTRFrmConvPos4 )
      Coil( #qOTSToNext )
   END_RUNG
   // the same network as SCL:
   #qOTSToNext := #sStWtRTRFrmConvPos4;
END_REGION

REGION Network 75: Transition for STATE Num:285 StL1S2Down
   RUNG wire#powerrail
      Contact( #sStL1S2Down )
      I_Contact( #sStWtResetRel )
      Contact( #sSst )
      Contact( #iL1S2Down )
      Coil( #sStL1S2Down_T1 )
   END_RUNG
   // the same network as SCL:
   #sStL1S2Down_T1 := #sStL1S2Down AND NOT #sStWtResetRel AND #sSst AND #iL1S2Down;
END_REGION

REGION Network 76: STATE Num:285 StL1S2Down
   RUNG wire#powerrail
      Contact( #sStL1S2Down )
      wire#w1
      I_Contact( #sStWtResetRel )
      I_Contact( #sStL1S2Down_T1 )
      wire#w2
      Coil( #sStL1S2Down )
   END_RUNG
   RUNG wire#powerrail
      Contact( #sStWtRTRFrmConvPos4_T1 )
   END_RUNG wire#w1
   RUNG wire#w2
      { S7_GenerateENO := "TRUE" } Move(in := 285, out1 => #StateNo)
   END_RUNG
   // the same network as SCL:
   #sStL1S2Down := (#sStL1S2Down OR #sStWtRTRFrmConvPos4_T1) AND NOT #sStWtResetRel AND NOT #sStL1S2Down_T1;
   IF #sStL1S2Down THEN #StateNo := 285; END_IF;
END_REGION

REGION Network 77: Actions for STATE Num:285 StL1S2Down
   RUNG wire#powerrail
      Contact( #sStL1S2Down )
      Coil( #qL1S2Down )
   END_RUNG
   // the same network as SCL:
   #qL1S2Down := #sStL1S2Down;
END_REGION

REGION Network 78: Transition for STATE Num:290 StWtL1TransBeginPos4
   RUNG wire#powerrail
      Contact( #sStWtL1TransBeginPos4 )
      I_Contact( #sStWtResetRel )
      Contact( #sSst )
      I_Contact( #iTransAreaClr )
      Coil( #sStWtL1TransBeginPos4_T1 )
   END_RUNG
   // the same network as SCL:
   #sStWtL1TransBeginPos4_T1 := #sStWtL1TransBeginPos4 AND NOT #sStWtResetRel AND #sSst AND NOT #iTransAreaClr;
END_REGION

REGION Network 79: STATE Num:290 StWtL1TransBeginPos4
   RUNG wire#powerrail
      Contact( #sStWtL1TransBeginPos4 )
      wire#w1
      I_Contact( #sStWtResetRel )
      I_Contact( #sStWtL1TransBeginPos4_T1 )
      wire#w2
      Coil( #sStWtL1TransBeginPos4 )
   END_RUNG
   RUNG wire#powerrail
      Contact( #sStL1S2Down_T1 )
   END_RUNG wire#w1
   RUNG wire#w2
      { S7_GenerateENO := "TRUE" } Move(in := 290, out1 => #StateNo)
   END_RUNG
   // the same network as SCL:
   #sStWtL1TransBeginPos4 := (#sStWtL1TransBeginPos4 OR #sStL1S2Down_T1) AND NOT #sStWtResetRel AND NOT #sStWtL1TransBeginPos4_T1;
   IF #sStWtL1TransBeginPos4 THEN #StateNo := 290; END_IF;
END_REGION

REGION Network 80: Transition for STATE Num:300 StWtTransDonePos4
   RUNG wire#powerrail
      Contact( #sStWtTransDonePos4 )
      I_Contact( #sStWtResetRel )
      Contact( #sSst )
      I_Contact( #iPalletPrsntL1 )
      Contact( #iTransAreaClr )
      Coil( #sStWtTransDonePos4_T1 )
   END_RUNG
   // the same network as SCL:
   #sStWtTransDonePos4_T1 := #sStWtTransDonePos4 AND NOT #sStWtResetRel AND #sSst AND NOT #iPalletPrsntL1 AND #iTransAreaClr;
END_REGION

REGION Network 81: STATE Num:300 StWtTransDonePos4
   RUNG wire#powerrail
      Contact( #sStWtTransDonePos4 )
      wire#w1
      I_Contact( #sStWtResetRel )
      I_Contact( #sStWtTransDonePos4_T1 )
      wire#w2
      Coil( #sStWtTransDonePos4 )
   END_RUNG
   RUNG wire#powerrail
      Contact( #sStWtL1TransBeginPos4_T1 )
   END_RUNG wire#w1
   RUNG wire#w2
      { S7_GenerateENO := "TRUE" } Move(in := 300, out1 => #StateNo)
   END_RUNG
   // the same network as SCL:
   #sStWtTransDonePos4 := (#sStWtTransDonePos4 OR #sStWtL1TransBeginPos4_T1) AND NOT #sStWtResetRel AND NOT #sStWtTransDonePos4_T1;
   IF #sStWtTransDonePos4 THEN #StateNo := 300; END_IF;
END_REGION

REGION Network 82: Transition for STATE Num:310 StChkPalletAtTT1
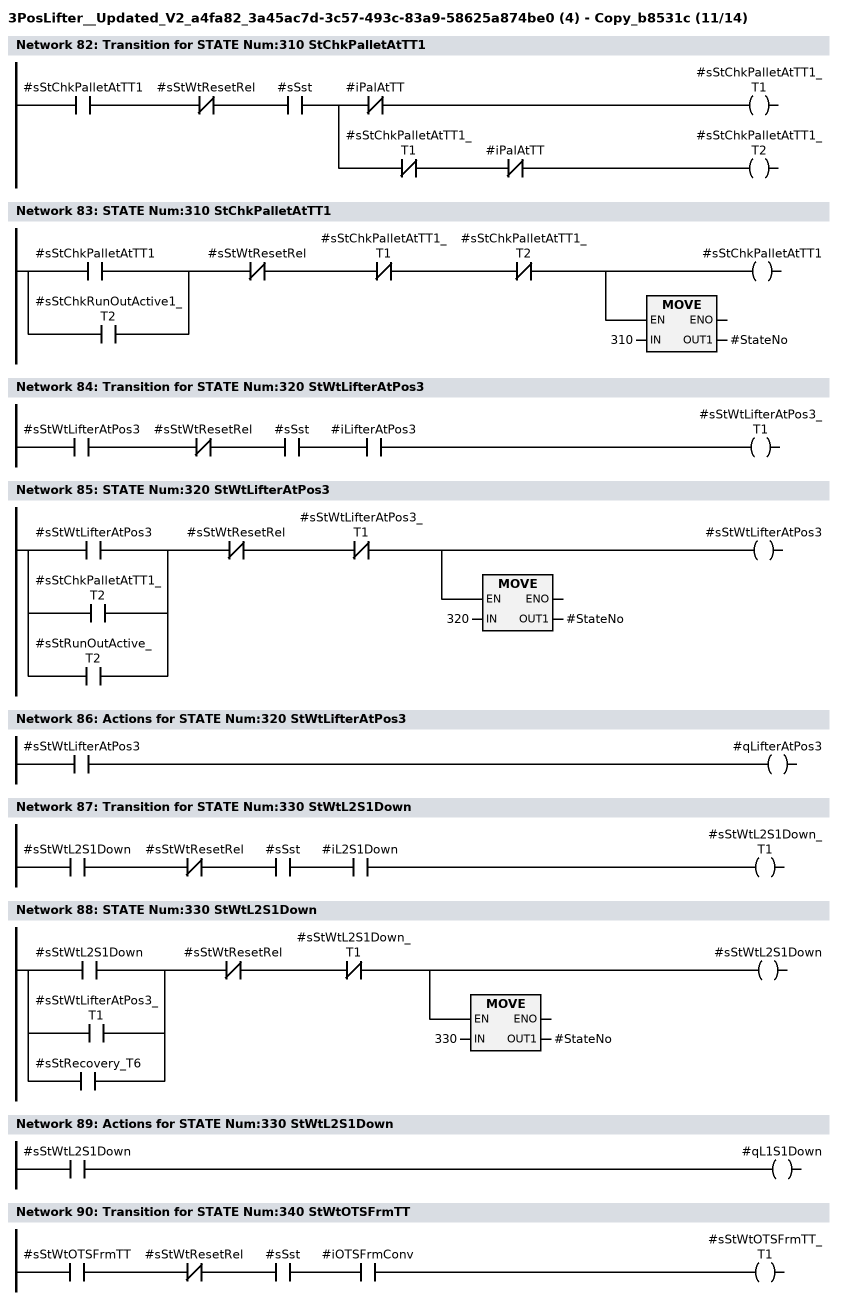
   RUNG wire#powerrail
      Contact( #sStChkPalletAtTT1 )
      I_Contact( #sStWtResetRel )
      Contact( #sSst )
      wire#w1
      I_Contact( #iPalAtTT )
      Coil( #sStChkPalletAtTT1_T1 )
   END_RUNG
   RUNG wire#w1
      I_Contact( #sStChkPalletAtTT1_T1 )
      I_Contact( #iPalAtTT )
      Coil( #sStChkPalletAtTT1_T2 )
   END_RUNG
   // the same network as SCL:
   #_w1 := #sStChkPalletAtTT1 AND NOT #sStWtResetRel AND #sSst;
   #sStChkPalletAtTT1_T1 := #_w1 AND NOT #iPalAtTT;
   #sStChkPalletAtTT1_T2 := #_w1 AND NOT #sStChkPalletAtTT1_T1 AND NOT #iPalAtTT;
END_REGION

REGION Network 83: STATE Num:310 StChkPalletAtTT1
   RUNG wire#powerrail
      Contact( #sStChkPalletAtTT1 )
      wire#w1
      I_Contact( #sStWtResetRel )
      I_Contact( #sStChkPalletAtTT1_T1 )
      I_Contact( #sStChkPalletAtTT1_T2 )
      wire#w2
      Coil( #sStChkPalletAtTT1 )
   END_RUNG
   RUNG wire#powerrail
      Contact( #sStChkRunOutActive1_T2 )
   END_RUNG wire#w1
   RUNG wire#w2
      { S7_GenerateENO := "TRUE" } Move(in := 310, out1 => #StateNo)
   END_RUNG
   // the same network as SCL:
   #sStChkPalletAtTT1 := (#sStChkPalletAtTT1 OR #sStChkRunOutActive1_T2) AND NOT #sStWtResetRel AND NOT #sStChkPalletAtTT1_T1 AND NOT #sStChkPalletAtTT1_T2;
   IF #sStChkPalletAtTT1 THEN #StateNo := 310; END_IF;
END_REGION

REGION Network 84: Transition for STATE Num:320 StWtLifterAtPos3
   RUNG wire#powerrail
      Contact( #sStWtLifterAtPos3 )
      I_Contact( #sStWtResetRel )
      Contact( #sSst )
      Contact( #iLifterAtPos3 )
      Coil( #sStWtLifterAtPos3_T1 )
   END_RUNG
   // the same network as SCL:
   #sStWtLifterAtPos3_T1 := #sStWtLifterAtPos3 AND NOT #sStWtResetRel AND #sSst AND #iLifterAtPos3;
END_REGION

REGION Network 85: STATE Num:320 StWtLifterAtPos3
   RUNG wire#powerrail
      Contact( #sStWtLifterAtPos3 )
      wire#w1
      I_Contact( #sStWtResetRel )
      I_Contact( #sStWtLifterAtPos3_T1 )
      wire#w2
      Coil( #sStWtLifterAtPos3 )
   END_RUNG
   RUNG wire#powerrail
      Contact( #sStChkPalletAtTT1_T2 )
   END_RUNG wire#w1
   RUNG wire#powerrail
      Contact( #sStRunOutActive_T2 )
   END_RUNG wire#w1
   RUNG wire#w2
      { S7_GenerateENO := "TRUE" } Move(in := 320, out1 => #StateNo)
   END_RUNG
   // the same network as SCL:
   #sStWtLifterAtPos3 := (#sStWtLifterAtPos3 OR #sStChkPalletAtTT1_T2 OR #sStRunOutActive_T2) AND NOT #sStWtResetRel AND NOT #sStWtLifterAtPos3_T1;
   IF #sStWtLifterAtPos3 THEN #StateNo := 320; END_IF;
END_REGION

REGION Network 86: Actions for STATE Num:320 StWtLifterAtPos3
   RUNG wire#powerrail
      Contact( #sStWtLifterAtPos3 )
      Coil( #qLifterAtPos3 )
   END_RUNG
   // the same network as SCL:
   #qLifterAtPos3 := #sStWtLifterAtPos3;
END_REGION

REGION Network 87: Transition for STATE Num:330 StWtL2S1Down
   RUNG wire#powerrail
      Contact( #sStWtL2S1Down )
      I_Contact( #sStWtResetRel )
      Contact( #sSst )
      Contact( #iL2S1Down )
      Coil( #sStWtL2S1Down_T1 )
   END_RUNG
   // the same network as SCL:
   #sStWtL2S1Down_T1 := #sStWtL2S1Down AND NOT #sStWtResetRel AND #sSst AND #iL2S1Down;
END_REGION

REGION Network 88: STATE Num:330 StWtL2S1Down
   RUNG wire#powerrail
      Contact( #sStWtL2S1Down )
      wire#w1
      I_Contact( #sStWtResetRel )
      I_Contact( #sStWtL2S1Down_T1 )
      wire#w2
      Coil( #sStWtL2S1Down )
   END_RUNG
   RUNG wire#powerrail
      Contact( #sStWtLifterAtPos3_T1 )
   END_RUNG wire#w1
   RUNG wire#powerrail
      Contact( #sStRecovery_T6 )
   END_RUNG wire#w1
   RUNG wire#w2
      { S7_GenerateENO := "TRUE" } Move(in := 330, out1 => #StateNo)
   END_RUNG
   // the same network as SCL:
   #sStWtL2S1Down := (#sStWtL2S1Down OR #sStWtLifterAtPos3_T1 OR #sStRecovery_T6) AND NOT #sStWtResetRel AND NOT #sStWtL2S1Down_T1;
   IF #sStWtL2S1Down THEN #StateNo := 330; END_IF;
END_REGION

REGION Network 89: Actions for STATE Num:330 StWtL2S1Down
   RUNG wire#powerrail
      Contact( #sStWtL2S1Down )
      Coil( #qL1S1Down )
   END_RUNG
   // the same network as SCL:
   #qL1S1Down := #sStWtL2S1Down;
END_REGION

REGION Network 90: Transition for STATE Num:340 StWtOTSFrmTT
   RUNG wire#powerrail
      Contact( #sStWtOTSFrmTT )
      I_Contact( #sStWtResetRel )
      Contact( #sSst )
      Contact( #iOTSFrmConv )
      Coil( #sStWtOTSFrmTT_T1 )
   END_RUNG
   // the same network as SCL:
   #sStWtOTSFrmTT_T1 := #sStWtOTSFrmTT AND NOT #sStWtResetRel AND #sSst AND #iOTSFrmConv;
END_REGION

REGION Network 91: STATE Num:340 StWtOTSFrmTT
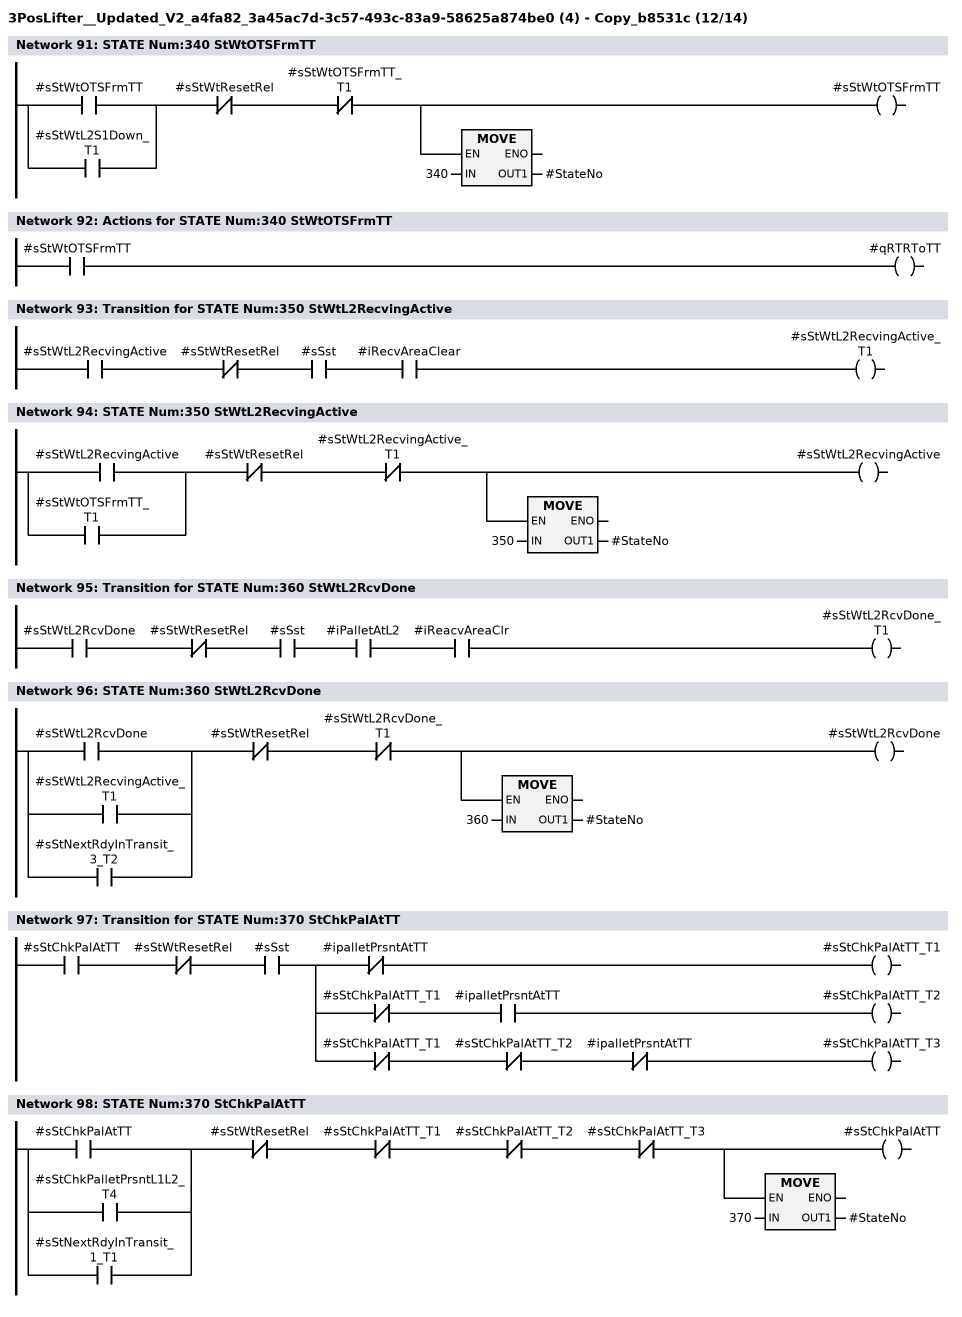
   RUNG wire#powerrail
      Contact( #sStWtOTSFrmTT )
      wire#w1
      I_Contact( #sStWtResetRel )
      I_Contact( #sStWtOTSFrmTT_T1 )
      wire#w2
      Coil( #sStWtOTSFrmTT )
   END_RUNG
   RUNG wire#powerrail
      Contact( #sStWtL2S1Down_T1 )
   END_RUNG wire#w1
   RUNG wire#w2
      { S7_GenerateENO := "TRUE" } Move(in := 340, out1 => #StateNo)
   END_RUNG
   // the same network as SCL:
   #sStWtOTSFrmTT := (#sStWtOTSFrmTT OR #sStWtL2S1Down_T1) AND NOT #sStWtResetRel AND NOT #sStWtOTSFrmTT_T1;
   IF #sStWtOTSFrmTT THEN #StateNo := 340; END_IF;
END_REGION

REGION Network 92: Actions for STATE Num:340 StWtOTSFrmTT
   RUNG wire#powerrail
      Contact( #sStWtOTSFrmTT )
      Coil( #qRTRToTT )
   END_RUNG
   // the same network as SCL:
   #qRTRToTT := #sStWtOTSFrmTT;
END_REGION

REGION Network 93: Transition for STATE Num:350 StWtL2RecvingActive
   RUNG wire#powerrail
      Contact( #sStWtL2RecvingActive )
      I_Contact( #sStWtResetRel )
      Contact( #sSst )
      Contact( #iRecvAreaClear )
      Coil( #sStWtL2RecvingActive_T1 )
   END_RUNG
   // the same network as SCL:
   #sStWtL2RecvingActive_T1 := #sStWtL2RecvingActive AND NOT #sStWtResetRel AND #sSst AND #iRecvAreaClear;
END_REGION

REGION Network 94: STATE Num:350 StWtL2RecvingActive
   RUNG wire#powerrail
      Contact( #sStWtL2RecvingActive )
      wire#w1
      I_Contact( #sStWtResetRel )
      I_Contact( #sStWtL2RecvingActive_T1 )
      wire#w2
      Coil( #sStWtL2RecvingActive )
   END_RUNG
   RUNG wire#powerrail
      Contact( #sStWtOTSFrmTT_T1 )
   END_RUNG wire#w1
   RUNG wire#w2
      { S7_GenerateENO := "TRUE" } Move(in := 350, out1 => #StateNo)
   END_RUNG
   // the same network as SCL:
   #sStWtL2RecvingActive := (#sStWtL2RecvingActive OR #sStWtOTSFrmTT_T1) AND NOT #sStWtResetRel AND NOT #sStWtL2RecvingActive_T1;
   IF #sStWtL2RecvingActive THEN #StateNo := 350; END_IF;
END_REGION

REGION Network 95: Transition for STATE Num:360 StWtL2RcvDone
   RUNG wire#powerrail
      Contact( #sStWtL2RcvDone )
      I_Contact( #sStWtResetRel )
      Contact( #sSst )
      Contact( #iPalletAtL2 )
      Contact( #iReacvAreaClr )
      Coil( #sStWtL2RcvDone_T1 )
   END_RUNG
   // the same network as SCL:
   #sStWtL2RcvDone_T1 := #sStWtL2RcvDone AND NOT #sStWtResetRel AND #sSst AND #iPalletAtL2 AND #iReacvAreaClr;
END_REGION

REGION Network 96: STATE Num:360 StWtL2RcvDone
   RUNG wire#powerrail
      Contact( #sStWtL2RcvDone )
      wire#w1
      I_Contact( #sStWtResetRel )
      I_Contact( #sStWtL2RcvDone_T1 )
      wire#w2
      Coil( #sStWtL2RcvDone )
   END_RUNG
   RUNG wire#powerrail
      Contact( #sStWtL2RecvingActive_T1 )
   END_RUNG wire#w1
   RUNG wire#powerrail
      Contact( #sStNextRdyInTransit_3_T2 )
   END_RUNG wire#w1
   RUNG wire#w2
      { S7_GenerateENO := "TRUE" } Move(in := 360, out1 => #StateNo)
   END_RUNG
   // the same network as SCL:
   #sStWtL2RcvDone := (#sStWtL2RcvDone OR #sStWtL2RecvingActive_T1 OR #sStNextRdyInTransit_3_T2) AND NOT #sStWtResetRel AND NOT #sStWtL2RcvDone_T1;
   IF #sStWtL2RcvDone THEN #StateNo := 360; END_IF;
END_REGION

REGION Network 97: Transition for STATE Num:370 StChkPalAtTT
   RUNG wire#powerrail
      Contact( #sStChkPalAtTT )
      I_Contact( #sStWtResetRel )
      Contact( #sSst )
      wire#w1
      I_Contact( #ipalletPrsntAtTT )
      Coil( #sStChkPalAtTT_T1 )
   END_RUNG
   RUNG wire#w1
      I_Contact( #sStChkPalAtTT_T1 )
      Contact( #ipalletPrsntAtTT )
      Coil( #sStChkPalAtTT_T2 )
   END_RUNG
   RUNG wire#w1
      I_Contact( #sStChkPalAtTT_T1 )
      I_Contact( #sStChkPalAtTT_T2 )
      I_Contact( #ipalletPrsntAtTT )
      Coil( #sStChkPalAtTT_T3 )
   END_RUNG
   // the same network as SCL:
   #_w1 := #sStChkPalAtTT AND NOT #sStWtResetRel AND #sSst;
   #sStChkPalAtTT_T1 := #_w1 AND NOT #ipalletPrsntAtTT;
   #sStChkPalAtTT_T2 := #_w1 AND NOT #sStChkPalAtTT_T1 AND #ipalletPrsntAtTT;
   #sStChkPalAtTT_T3 := #_w1 AND NOT #sStChkPalAtTT_T1 AND NOT #sStChkPalAtTT_T2 AND NOT #ipalletPrsntAtTT;
END_REGION

REGION Network 98: STATE Num:370 StChkPalAtTT
   RUNG wire#powerrail
      Contact( #sStChkPalAtTT )
      wire#w1
      I_Contact( #sStWtResetRel )
      I_Contact( #sStChkPalAtTT_T1 )
      I_Contact( #sStChkPalAtTT_T2 )
      I_Contact( #sStChkPalAtTT_T3 )
      wire#w2
      Coil( #sStChkPalAtTT )
   END_RUNG
   RUNG wire#powerrail
      Contact( #sStChkPalletPrsntL1L2_T4 )
   END_RUNG wire#w1
   RUNG wire#powerrail
      Contact( #sStNextRdyInTransit_1_T1 )
   END_RUNG wire#w1
   RUNG wire#w2
      { S7_GenerateENO := "TRUE" } Move(in := 370, out1 => #StateNo)
   END_RUNG
   // the same network as SCL:
   #sStChkPalAtTT := (#sStChkPalAtTT OR #sStChkPalletPrsntL1L2_T4 OR #sStNextRdyInTransit_1_T1) AND NOT #sStWtResetRel AND NOT #sStChkPalAtTT_T1 AND NOT #sStChkPalAtTT_T2 AND NOT #sStChkPalAtTT_T3;
   IF #sStChkPalAtTT THEN #StateNo := 370; END_IF;
END_REGION

REGION Network 99: Transition for STATE Num:380 StWtLifterAtPos2
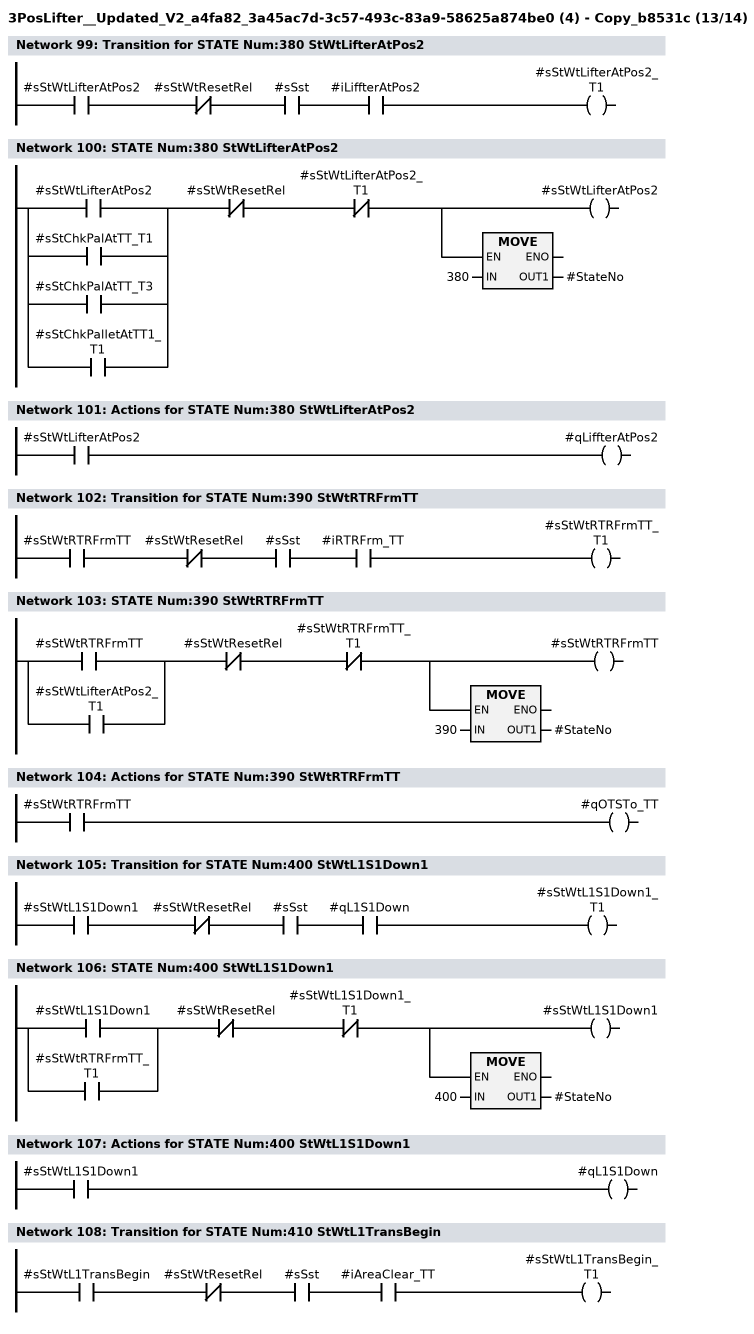
   RUNG wire#powerrail
      Contact( #sStWtLifterAtPos2 )
      I_Contact( #sStWtResetRel )
      Contact( #sSst )
      Contact( #iLiffterAtPos2 )
      Coil( #sStWtLifterAtPos2_T1 )
   END_RUNG
   // the same network as SCL:
   #sStWtLifterAtPos2_T1 := #sStWtLifterAtPos2 AND NOT #sStWtResetRel AND #sSst AND #iLiffterAtPos2;
END_REGION

REGION Network 100: STATE Num:380 StWtLifterAtPos2
   RUNG wire#powerrail
      Contact( #sStWtLifterAtPos2 )
      wire#w1
      I_Contact( #sStWtResetRel )
      I_Contact( #sStWtLifterAtPos2_T1 )
      wire#w2
      Coil( #sStWtLifterAtPos2 )
   END_RUNG
   RUNG wire#powerrail
      Contact( #sStChkPalAtTT_T1 )
   END_RUNG wire#w1
   RUNG wire#powerrail
      Contact( #sStChkPalAtTT_T3 )
   END_RUNG wire#w1
   RUNG wire#powerrail
      Contact( #sStChkPalletAtTT1_T1 )
   END_RUNG wire#w1
   RUNG wire#w2
      { S7_GenerateENO := "TRUE" } Move(in := 380, out1 => #StateNo)
   END_RUNG
   // the same network as SCL:
   #sStWtLifterAtPos2 := (#sStWtLifterAtPos2 OR #sStChkPalAtTT_T1 OR #sStChkPalAtTT_T3 OR #sStChkPalletAtTT1_T1) AND NOT #sStWtResetRel AND NOT #sStWtLifterAtPos2_T1;
   IF #sStWtLifterAtPos2 THEN #StateNo := 380; END_IF;
END_REGION

REGION Network 101: Actions for STATE Num:380 StWtLifterAtPos2
   RUNG wire#powerrail
      Contact( #sStWtLifterAtPos2 )
      Coil( #qLiffterAtPos2 )
   END_RUNG
   // the same network as SCL:
   #qLiffterAtPos2 := #sStWtLifterAtPos2;
END_REGION

REGION Network 102: Transition for STATE Num:390 StWtRTRFrmTT
   RUNG wire#powerrail
      Contact( #sStWtRTRFrmTT )
      I_Contact( #sStWtResetRel )
      Contact( #sSst )
      Contact( #iRTRFrm_TT )
      Coil( #sStWtRTRFrmTT_T1 )
   END_RUNG
   // the same network as SCL:
   #sStWtRTRFrmTT_T1 := #sStWtRTRFrmTT AND NOT #sStWtResetRel AND #sSst AND #iRTRFrm_TT;
END_REGION

REGION Network 103: STATE Num:390 StWtRTRFrmTT
   RUNG wire#powerrail
      Contact( #sStWtRTRFrmTT )
      wire#w1
      I_Contact( #sStWtResetRel )
      I_Contact( #sStWtRTRFrmTT_T1 )
      wire#w2
      Coil( #sStWtRTRFrmTT )
   END_RUNG
   RUNG wire#powerrail
      Contact( #sStWtLifterAtPos2_T1 )
   END_RUNG wire#w1
   RUNG wire#w2
      { S7_GenerateENO := "TRUE" } Move(in := 390, out1 => #StateNo)
   END_RUNG
   // the same network as SCL:
   #sStWtRTRFrmTT := (#sStWtRTRFrmTT OR #sStWtLifterAtPos2_T1) AND NOT #sStWtResetRel AND NOT #sStWtRTRFrmTT_T1;
   IF #sStWtRTRFrmTT THEN #StateNo := 390; END_IF;
END_REGION

REGION Network 104: Actions for STATE Num:390 StWtRTRFrmTT
   RUNG wire#powerrail
      Contact( #sStWtRTRFrmTT )
      Coil( #qOTSTo_TT )
   END_RUNG
   // the same network as SCL:
   #qOTSTo_TT := #sStWtRTRFrmTT;
END_REGION

REGION Network 105: Transition for STATE Num:400 StWtL1S1Down1
   RUNG wire#powerrail
      Contact( #sStWtL1S1Down1 )
      I_Contact( #sStWtResetRel )
      Contact( #sSst )
      Contact( #qL1S1Down )
      Coil( #sStWtL1S1Down1_T1 )
   END_RUNG
   // the same network as SCL:
   #sStWtL1S1Down1_T1 := #sStWtL1S1Down1 AND NOT #sStWtResetRel AND #sSst AND #qL1S1Down;
END_REGION

REGION Network 106: STATE Num:400 StWtL1S1Down1
   RUNG wire#powerrail
      Contact( #sStWtL1S1Down1 )
      wire#w1
      I_Contact( #sStWtResetRel )
      I_Contact( #sStWtL1S1Down1_T1 )
      wire#w2
      Coil( #sStWtL1S1Down1 )
   END_RUNG
   RUNG wire#powerrail
      Contact( #sStWtRTRFrmTT_T1 )
   END_RUNG wire#w1
   RUNG wire#w2
      { S7_GenerateENO := "TRUE" } Move(in := 400, out1 => #StateNo)
   END_RUNG
   // the same network as SCL:
   #sStWtL1S1Down1 := (#sStWtL1S1Down1 OR #sStWtRTRFrmTT_T1) AND NOT #sStWtResetRel AND NOT #sStWtL1S1Down1_T1;
   IF #sStWtL1S1Down1 THEN #StateNo := 400; END_IF;
END_REGION

REGION Network 107: Actions for STATE Num:400 StWtL1S1Down1
   RUNG wire#powerrail
      Contact( #sStWtL1S1Down1 )
      Coil( #qL1S1Down )
   END_RUNG
   // the same network as SCL:
   #qL1S1Down := #sStWtL1S1Down1;
END_REGION

REGION Network 108: Transition for STATE Num:410 StWtL1TransBegin
   RUNG wire#powerrail
      Contact( #sStWtL1TransBegin )
      I_Contact( #sStWtResetRel )
      Contact( #sSst )
      Contact( #iAreaClear_TT )
      Coil( #sStWtL1TransBegin_T1 )
   END_RUNG
   // the same network as SCL:
   #sStWtL1TransBegin_T1 := #sStWtL1TransBegin AND NOT #sStWtResetRel AND #sSst AND #iAreaClear_TT;
END_REGION

REGION Network 109: STATE Num:410 StWtL1TransBegin
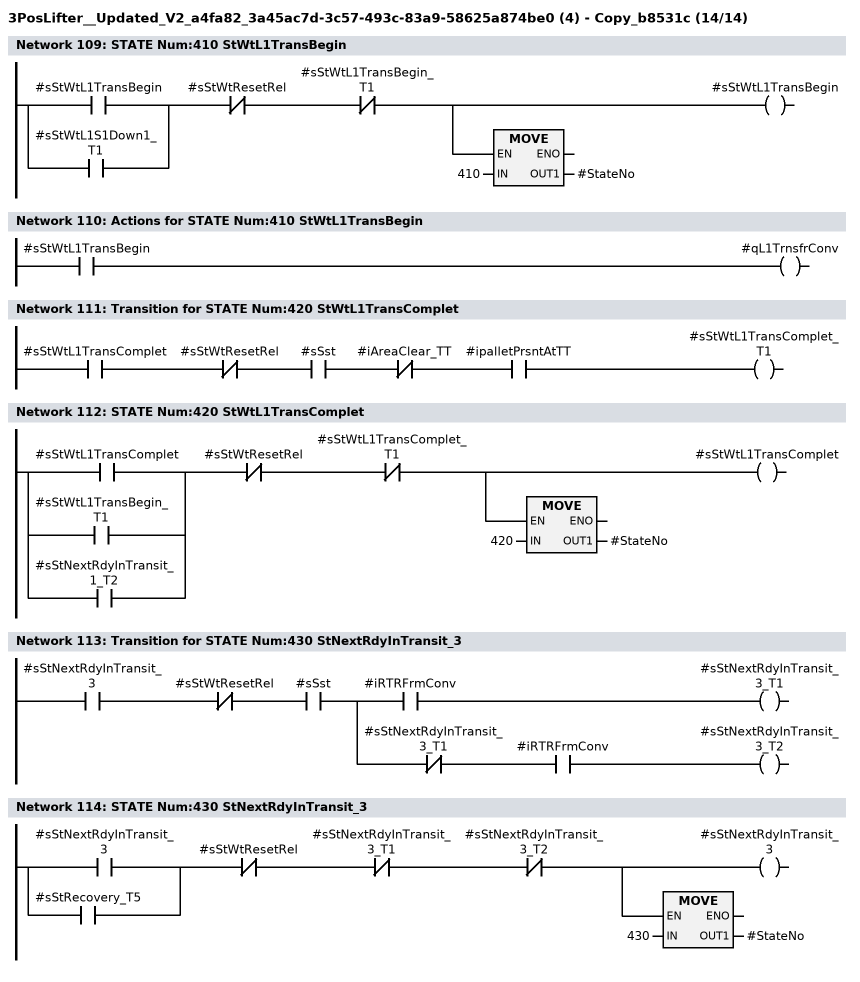
   RUNG wire#powerrail
      Contact( #sStWtL1TransBegin )
      wire#w1
      I_Contact( #sStWtResetRel )
      I_Contact( #sStWtL1TransBegin_T1 )
      wire#w2
      Coil( #sStWtL1TransBegin )
   END_RUNG
   RUNG wire#powerrail
      Contact( #sStWtL1S1Down1_T1 )
   END_RUNG wire#w1
   RUNG wire#w2
      { S7_GenerateENO := "TRUE" } Move(in := 410, out1 => #StateNo)
   END_RUNG
   // the same network as SCL:
   #sStWtL1TransBegin := (#sStWtL1TransBegin OR #sStWtL1S1Down1_T1) AND NOT #sStWtResetRel AND NOT #sStWtL1TransBegin_T1;
   IF #sStWtL1TransBegin THEN #StateNo := 410; END_IF;
END_REGION

REGION Network 110: Actions for STATE Num:410 StWtL1TransBegin
   RUNG wire#powerrail
      Contact( #sStWtL1TransBegin )
      Coil( #qL1TrnsfrConv )
   END_RUNG
   // the same network as SCL:
   #qL1TrnsfrConv := #sStWtL1TransBegin;
END_REGION

REGION Network 111: Transition for STATE Num:420 StWtL1TransComplet
   RUNG wire#powerrail
      Contact( #sStWtL1TransComplet )
      I_Contact( #sStWtResetRel )
      Contact( #sSst )
      I_Contact( #iAreaClear_TT )
      Contact( #ipalletPrsntAtTT )
      Coil( #sStWtL1TransComplet_T1 )
   END_RUNG
   // the same network as SCL:
   #sStWtL1TransComplet_T1 := #sStWtL1TransComplet AND NOT #sStWtResetRel AND #sSst AND NOT #iAreaClear_TT AND #ipalletPrsntAtTT;
END_REGION

REGION Network 112: STATE Num:420 StWtL1TransComplet
   RUNG wire#powerrail
      Contact( #sStWtL1TransComplet )
      wire#w1
      I_Contact( #sStWtResetRel )
      I_Contact( #sStWtL1TransComplet_T1 )
      wire#w2
      Coil( #sStWtL1TransComplet )
   END_RUNG
   RUNG wire#powerrail
      Contact( #sStWtL1TransBegin_T1 )
   END_RUNG wire#w1
   RUNG wire#powerrail
      Contact( #sStNextRdyInTransit_1_T2 )
   END_RUNG wire#w1
   RUNG wire#w2
      { S7_GenerateENO := "TRUE" } Move(in := 420, out1 => #StateNo)
   END_RUNG
   // the same network as SCL:
   #sStWtL1TransComplet := (#sStWtL1TransComplet OR #sStWtL1TransBegin_T1 OR #sStNextRdyInTransit_1_T2) AND NOT #sStWtResetRel AND NOT #sStWtL1TransComplet_T1;
   IF #sStWtL1TransComplet THEN #StateNo := 420; END_IF;
END_REGION

REGION Network 113: Transition for STATE Num:430 StNextRdyInTransit_3
   RUNG wire#powerrail
      Contact( #sStNextRdyInTransit_3 )
      I_Contact( #sStWtResetRel )
      Contact( #sSst )
      wire#w1
      Contact( #iRTRFrmConv )
      Coil( #sStNextRdyInTransit_3_T1 )
   END_RUNG
   RUNG wire#w1
      I_Contact( #sStNextRdyInTransit_3_T1 )
      Contact( #iRTRFrmConv )
      Coil( #sStNextRdyInTransit_3_T2 )
   END_RUNG
   // the same network as SCL:
   #_w1 := #sStNextRdyInTransit_3 AND NOT #sStWtResetRel AND #sSst;
   #sStNextRdyInTransit_3_T1 := #_w1 AND #iRTRFrmConv;
   #sStNextRdyInTransit_3_T2 := #_w1 AND NOT #sStNextRdyInTransit_3_T1 AND #iRTRFrmConv;
END_REGION

REGION Network 114: STATE Num:430 StNextRdyInTransit_3
   RUNG wire#powerrail
      Contact( #sStNextRdyInTransit_3 )
      wire#w1
      I_Contact( #sStWtResetRel )
      I_Contact( #sStNextRdyInTransit_3_T1 )
      I_Contact( #sStNextRdyInTransit_3_T2 )
      wire#w2
      Coil( #sStNextRdyInTransit_3 )
   END_RUNG
   RUNG wire#powerrail
      Contact( #sStRecovery_T5 )
   END_RUNG wire#w1
   RUNG wire#w2
      { S7_GenerateENO := "TRUE" } Move(in := 430, out1 => #StateNo)
   END_RUNG
   // the same network as SCL:
   #sStNextRdyInTransit_3 := (#sStNextRdyInTransit_3 OR #sStRecovery_T5) AND NOT #sStWtResetRel AND NOT #sStNextRdyInTransit_3_T1 AND NOT #sStNextRdyInTransit_3_T2;
   IF #sStNextRdyInTransit_3 THEN #StateNo := 430; END_IF;
END_REGION
END_FUNCTION_BLOCK

FUNCTION_BLOCK "FB_CentreStand_Fix_Seq"   // FB1, LAD
VERSION : 0.1
// stored: AutoNumber true, IsIECCheckEnabled false, UDAEnableTagReadback false
   VAR_INPUT
      iAutoRunning : Bool;
      iFixClamp : Bool;
      iFixEmpty : Bool;
      iFixTrayPresent : Bool;
      iFixUnclamp : Bool;
      iR1DropOver : Bool;
      iR1PickOver : Bool;
      iR2OperationOver : Bool;
      iR2ServiceActivated : Bool;
      iReset_fault : Bool;
      iRobotOutofZone : Bool;
      iSstMode : Bool;
      iSstPB : Bool;
   END_VAR
   VAR_OUTPUT
      qFixClamp : Bool;
      qFixUnclamp : Bool;
      qR1ReadytoDropTray : Bool;
      qR1ReadytoPickTray : Bool;
      qR2OperationStart : Bool;
   END_VAR
   VAR_IN_OUT
      iqR2ServiceActive : Bool;
      iqR2ServiceCompleted : Bool;
   END_VAR
   VAR DB_SPECIFIC
      StateNo : Int;
      s138_WaitBothRbtOutAl : Bool;
      s138_WaitBothRbtOutAl_T1 : Bool;
      s138_WaitBothRbtOutAl_T2 : Bool;
      s139_FixEmpty : Bool;
      s139_FixEmpty_T1 : Bool;
      s140_FixTrayPrsntRec : Bool;
      s140_FixTrayPrsntRec_T1 : Bool;
      s140_FixTrayPrsntRec_T2 : Bool;
      s141_FixUnclampCmd : Bool;
      s141_FixUnclampCmd_T1 : Bool;
      s142_TrayRdyDropFix : Bool;
      s142_TrayRdyDropFix_T1 : Bool;
      s143_RbtDropFixChkTr : Bool;
      s143_RbtDropFixChkTr_T1 : Bool;
      s144_RbtOutAreaDrop : Bool;
      s144_RbtOutAreaDrop_T1 : Bool;
      s145_FixClamp : Bool;
      s145_FixClamp_T1 : Bool;
      s146_Rbt2AlloyOpOver : Bool;
      s146_Rbt2AlloyOpOver_T1 : Bool;
      s147_FixUnclmpCmdAft : Bool;
      s147_FixUnclmpCmdAft_T1 : Bool;
      s148_RdyPickTrayAftr : Bool;
      s148_RdyPickTrayAftr_T1 : Bool;
      s149_RbtPickTrayChkE : Bool;
      s149_RbtPickTrayChkE_T1 : Bool;
      s191_WaitRbt2OutArea : Bool;
      s191_WaitRbt2OutArea_T1 : Bool;
      sSst : Bool;
      sSstPulse : Bool;
      sSstRise : Bool;
      sStWtResetRel : Bool;
      sStWtResetRel_T1 : Bool;
   END_VAR
   VAR_TEMP
      c138_WaitBothRbtOutAl_T1 : Bool;
      c138_WaitBothRbtOutAl_T2 : Bool;
      c140_FixTrayPrsntRec_T1 : Bool;
      c140_FixTrayPrsntRec_T2 : Bool;
      tOne : Bool;
   END_VAR
   VAR_TEMP   // added for the SCL form of the ladder/FBD networks
      _w1 : Bool;
   END_VAR
BEGIN

REGION Network 1
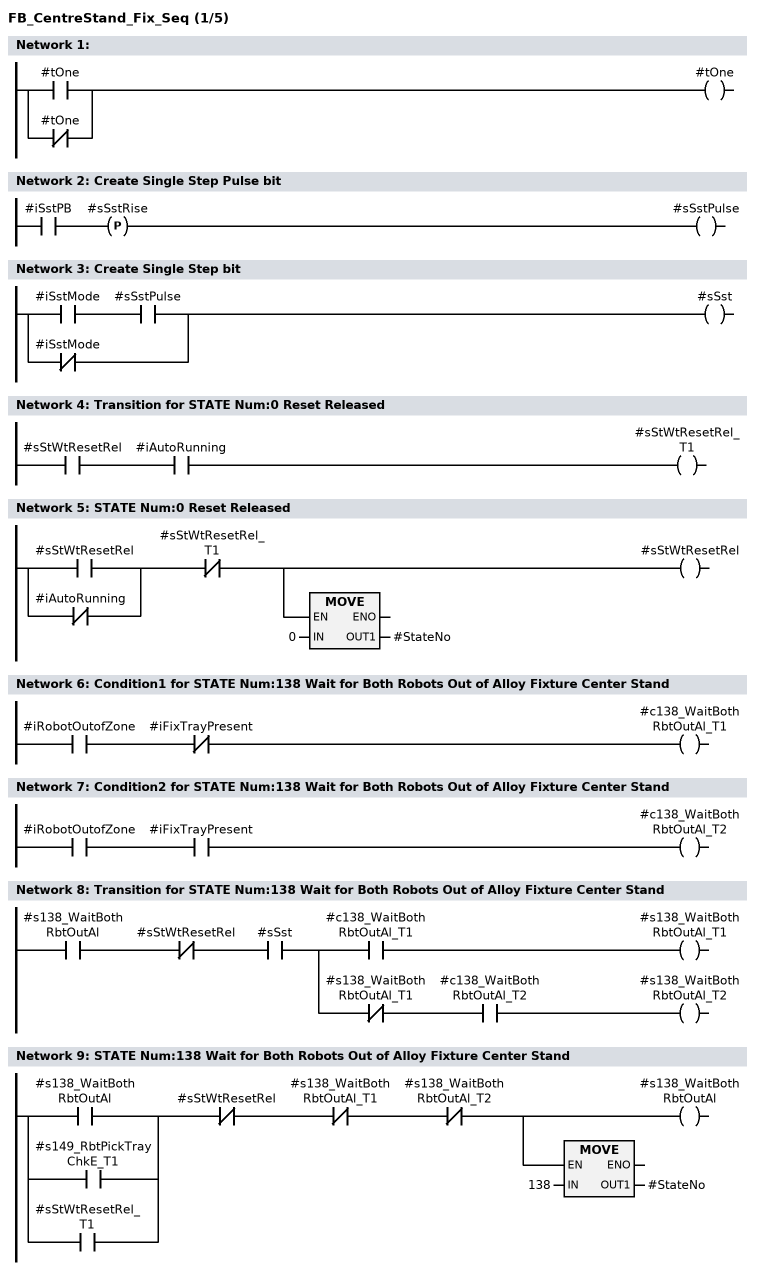
   RUNG wire#powerrail
      Contact( #tOne )
      wire#w1
      Coil( #tOne )
   END_RUNG
   RUNG wire#powerrail
      I_Contact( #tOne )
   END_RUNG wire#w1
   // the same network as SCL:
   #tOne := #tOne OR NOT #tOne;
END_REGION

REGION Network 2: Create Single Step Pulse bit
   RUNG wire#powerrail
      Contact( #iSstPB )
      P_Trig( #sSstRise )
      Coil( #sSstPulse )
   END_RUNG
   // the same network as SCL:
   #_w1 := #iSstPB AND NOT #sSstRise;   // rising edge
   #sSstRise := #iSstPB;
   #sSstPulse := #_w1;
END_REGION

REGION Network 3: Create Single Step bit
   RUNG wire#powerrail
      Contact( #iSstMode )
      Contact( #sSstPulse )
      wire#w1
      Coil( #sSst )
   END_RUNG
   RUNG wire#powerrail
      I_Contact( #iSstMode )
   END_RUNG wire#w1
   // the same network as SCL:
   #sSst := (#iSstMode AND #sSstPulse) OR NOT #iSstMode;
END_REGION

REGION Network 4: Transition for STATE Num:0 Reset Released
   RUNG wire#powerrail
      Contact( #sStWtResetRel )
      Contact( #iAutoRunning )
      Coil( #sStWtResetRel_T1 )
   END_RUNG
   // the same network as SCL:
   #sStWtResetRel_T1 := #sStWtResetRel AND #iAutoRunning;
END_REGION

REGION Network 5: STATE Num:0 Reset Released
   RUNG wire#powerrail
      Contact( #sStWtResetRel )
      wire#w1
      I_Contact( #sStWtResetRel_T1 )
      wire#w2
      Coil( #sStWtResetRel )
   END_RUNG
   RUNG wire#powerrail
      I_Contact( #iAutoRunning )
   END_RUNG wire#w1
   RUNG wire#w2
      { S7_GenerateENO := "TRUE" } Move(in := 0, out1 => #StateNo)
   END_RUNG
   // the same network as SCL:
   #sStWtResetRel := (#sStWtResetRel OR NOT #iAutoRunning) AND NOT #sStWtResetRel_T1;
   IF #sStWtResetRel THEN #StateNo := 0; END_IF;
END_REGION

REGION Network 6: Condition1 for STATE Num:138 Wait for Both Robots Out of Alloy Fixture Center Stand
   RUNG wire#powerrail
      Contact( #iRobotOutofZone )
      I_Contact( #iFixTrayPresent )
      Coil( #c138_WaitBothRbtOutAl_T1 )
   END_RUNG
   // the same network as SCL:
   #c138_WaitBothRbtOutAl_T1 := #iRobotOutofZone AND NOT #iFixTrayPresent;
END_REGION

REGION Network 7: Condition2 for STATE Num:138 Wait for Both Robots Out of Alloy Fixture Center Stand
   RUNG wire#powerrail
      Contact( #iRobotOutofZone )
      Contact( #iFixTrayPresent )
      Coil( #c138_WaitBothRbtOutAl_T2 )
   END_RUNG
   // the same network as SCL:
   #c138_WaitBothRbtOutAl_T2 := #iRobotOutofZone AND #iFixTrayPresent;
END_REGION

REGION Network 8: Transition for STATE Num:138 Wait for Both Robots Out of Alloy Fixture Center Stand
   RUNG wire#powerrail
      Contact( #s138_WaitBothRbtOutAl )
      I_Contact( #sStWtResetRel )
      Contact( #sSst )
      wire#w1
      Contact( #c138_WaitBothRbtOutAl_T1 )
      Coil( #s138_WaitBothRbtOutAl_T1 )
   END_RUNG
   RUNG wire#w1
      I_Contact( #s138_WaitBothRbtOutAl_T1 )
      Contact( #c138_WaitBothRbtOutAl_T2 )
      Coil( #s138_WaitBothRbtOutAl_T2 )
   END_RUNG
   // the same network as SCL:
   #_w1 := #s138_WaitBothRbtOutAl AND NOT #sStWtResetRel AND #sSst;
   #s138_WaitBothRbtOutAl_T1 := #_w1 AND #c138_WaitBothRbtOutAl_T1;
   #s138_WaitBothRbtOutAl_T2 := #_w1 AND NOT #s138_WaitBothRbtOutAl_T1 AND #c138_WaitBothRbtOutAl_T2;
END_REGION

REGION Network 9: STATE Num:138 Wait for Both Robots Out of Alloy Fixture Center Stand
   RUNG wire#powerrail
      Contact( #s138_WaitBothRbtOutAl )
      wire#w1
      I_Contact( #sStWtResetRel )
      I_Contact( #s138_WaitBothRbtOutAl_T1 )
      I_Contact( #s138_WaitBothRbtOutAl_T2 )
      wire#w2
      Coil( #s138_WaitBothRbtOutAl )
   END_RUNG
   RUNG wire#powerrail
      Contact( #s149_RbtPickTrayChkE_T1 )
   END_RUNG wire#w1
   RUNG wire#powerrail
      Contact( #sStWtResetRel_T1 )
   END_RUNG wire#w1
   RUNG wire#w2
      { S7_GenerateENO := "TRUE" } Move(in := 138, out1 => #StateNo)
   END_RUNG
   // the same network as SCL:
   #s138_WaitBothRbtOutAl := (#s138_WaitBothRbtOutAl OR #s149_RbtPickTrayChkE_T1 OR #sStWtResetRel_T1) AND NOT #sStWtResetRel AND NOT #s138_WaitBothRbtOutAl_T1 AND NOT #s138_WaitBothRbtOutAl_T2;
   IF #s138_WaitBothRbtOutAl THEN #StateNo := 138; END_IF;
END_REGION

REGION Network 10: Transition for STATE Num:139 Fix Empty
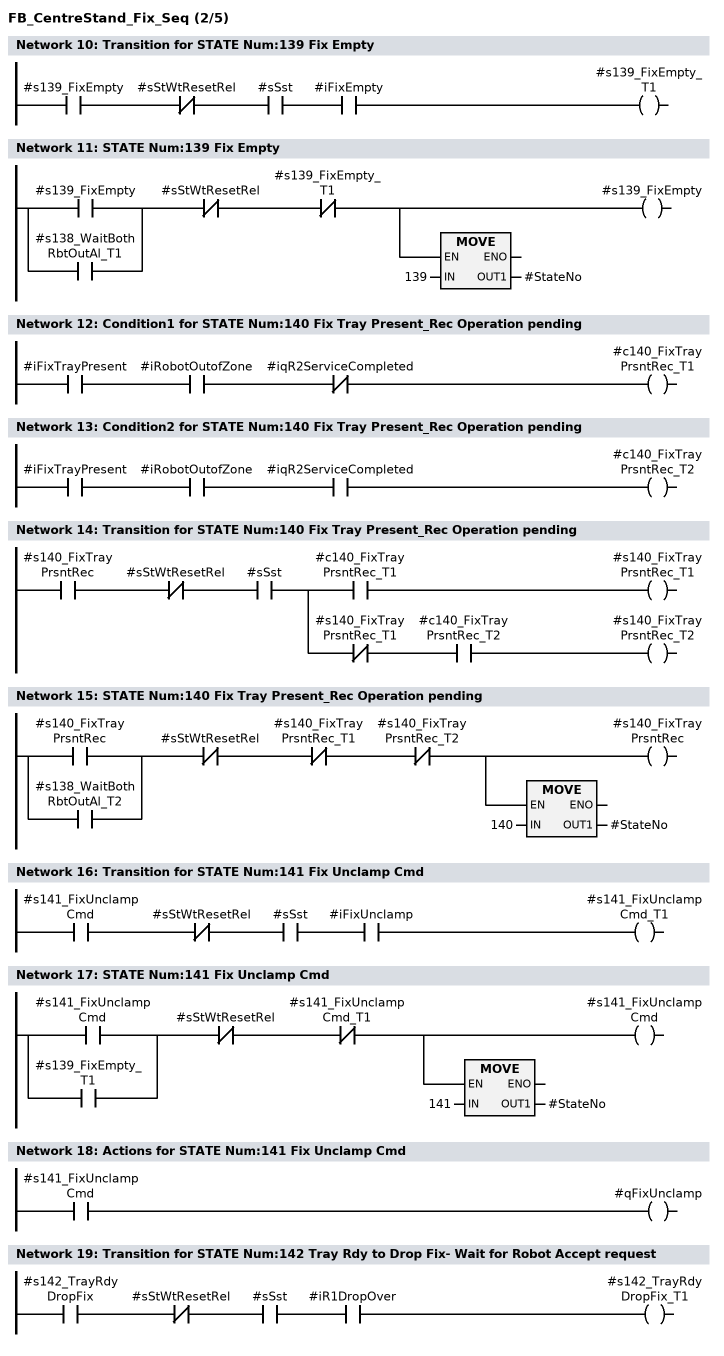
   RUNG wire#powerrail
      Contact( #s139_FixEmpty )
      I_Contact( #sStWtResetRel )
      Contact( #sSst )
      Contact( #iFixEmpty )
      Coil( #s139_FixEmpty_T1 )
   END_RUNG
   // the same network as SCL:
   #s139_FixEmpty_T1 := #s139_FixEmpty AND NOT #sStWtResetRel AND #sSst AND #iFixEmpty;
END_REGION

REGION Network 11: STATE Num:139 Fix Empty
   RUNG wire#powerrail
      Contact( #s139_FixEmpty )
      wire#w1
      I_Contact( #sStWtResetRel )
      I_Contact( #s139_FixEmpty_T1 )
      wire#w2
      Coil( #s139_FixEmpty )
   END_RUNG
   RUNG wire#powerrail
      Contact( #s138_WaitBothRbtOutAl_T1 )
   END_RUNG wire#w1
   RUNG wire#w2
      { S7_GenerateENO := "TRUE" } Move(in := 139, out1 => #StateNo)
   END_RUNG
   // the same network as SCL:
   #s139_FixEmpty := (#s139_FixEmpty OR #s138_WaitBothRbtOutAl_T1) AND NOT #sStWtResetRel AND NOT #s139_FixEmpty_T1;
   IF #s139_FixEmpty THEN #StateNo := 139; END_IF;
END_REGION

REGION Network 12: Condition1 for STATE Num:140 Fix Tray Present_Rec Operation pending
   RUNG wire#powerrail
      Contact( #iFixTrayPresent )
      Contact( #iRobotOutofZone )
      I_Contact( #iqR2ServiceCompleted )
      Coil( #c140_FixTrayPrsntRec_T1 )
   END_RUNG
   // the same network as SCL:
   #c140_FixTrayPrsntRec_T1 := #iFixTrayPresent AND #iRobotOutofZone AND NOT #iqR2ServiceCompleted;
END_REGION

REGION Network 13: Condition2 for STATE Num:140 Fix Tray Present_Rec Operation pending
   RUNG wire#powerrail
      Contact( #iFixTrayPresent )
      Contact( #iRobotOutofZone )
      Contact( #iqR2ServiceCompleted )
      Coil( #c140_FixTrayPrsntRec_T2 )
   END_RUNG
   // the same network as SCL:
   #c140_FixTrayPrsntRec_T2 := #iFixTrayPresent AND #iRobotOutofZone AND #iqR2ServiceCompleted;
END_REGION

REGION Network 14: Transition for STATE Num:140 Fix Tray Present_Rec Operation pending
   RUNG wire#powerrail
      Contact( #s140_FixTrayPrsntRec )
      I_Contact( #sStWtResetRel )
      Contact( #sSst )
      wire#w1
      Contact( #c140_FixTrayPrsntRec_T1 )
      Coil( #s140_FixTrayPrsntRec_T1 )
   END_RUNG
   RUNG wire#w1
      I_Contact( #s140_FixTrayPrsntRec_T1 )
      Contact( #c140_FixTrayPrsntRec_T2 )
      Coil( #s140_FixTrayPrsntRec_T2 )
   END_RUNG
   // the same network as SCL:
   #_w1 := #s140_FixTrayPrsntRec AND NOT #sStWtResetRel AND #sSst;
   #s140_FixTrayPrsntRec_T1 := #_w1 AND #c140_FixTrayPrsntRec_T1;
   #s140_FixTrayPrsntRec_T2 := #_w1 AND NOT #s140_FixTrayPrsntRec_T1 AND #c140_FixTrayPrsntRec_T2;
END_REGION

REGION Network 15: STATE Num:140 Fix Tray Present_Rec Operation pending
   RUNG wire#powerrail
      Contact( #s140_FixTrayPrsntRec )
      wire#w1
      I_Contact( #sStWtResetRel )
      I_Contact( #s140_FixTrayPrsntRec_T1 )
      I_Contact( #s140_FixTrayPrsntRec_T2 )
      wire#w2
      Coil( #s140_FixTrayPrsntRec )
   END_RUNG
   RUNG wire#powerrail
      Contact( #s138_WaitBothRbtOutAl_T2 )
   END_RUNG wire#w1
   RUNG wire#w2
      { S7_GenerateENO := "TRUE" } Move(in := 140, out1 => #StateNo)
   END_RUNG
   // the same network as SCL:
   #s140_FixTrayPrsntRec := (#s140_FixTrayPrsntRec OR #s138_WaitBothRbtOutAl_T2) AND NOT #sStWtResetRel AND NOT #s140_FixTrayPrsntRec_T1 AND NOT #s140_FixTrayPrsntRec_T2;
   IF #s140_FixTrayPrsntRec THEN #StateNo := 140; END_IF;
END_REGION

REGION Network 16: Transition for STATE Num:141 Fix Unclamp Cmd
   RUNG wire#powerrail
      Contact( #s141_FixUnclampCmd )
      I_Contact( #sStWtResetRel )
      Contact( #sSst )
      Contact( #iFixUnclamp )
      Coil( #s141_FixUnclampCmd_T1 )
   END_RUNG
   // the same network as SCL:
   #s141_FixUnclampCmd_T1 := #s141_FixUnclampCmd AND NOT #sStWtResetRel AND #sSst AND #iFixUnclamp;
END_REGION

REGION Network 17: STATE Num:141 Fix Unclamp Cmd
   RUNG wire#powerrail
      Contact( #s141_FixUnclampCmd )
      wire#w1
      I_Contact( #sStWtResetRel )
      I_Contact( #s141_FixUnclampCmd_T1 )
      wire#w2
      Coil( #s141_FixUnclampCmd )
   END_RUNG
   RUNG wire#powerrail
      Contact( #s139_FixEmpty_T1 )
   END_RUNG wire#w1
   RUNG wire#w2
      { S7_GenerateENO := "TRUE" } Move(in := 141, out1 => #StateNo)
   END_RUNG
   // the same network as SCL:
   #s141_FixUnclampCmd := (#s141_FixUnclampCmd OR #s139_FixEmpty_T1) AND NOT #sStWtResetRel AND NOT #s141_FixUnclampCmd_T1;
   IF #s141_FixUnclampCmd THEN #StateNo := 141; END_IF;
END_REGION

REGION Network 18: Actions for STATE Num:141 Fix Unclamp Cmd
   RUNG wire#powerrail
      Contact( #s141_FixUnclampCmd )
      Coil( #qFixUnclamp )
   END_RUNG
   // the same network as SCL:
   #qFixUnclamp := #s141_FixUnclampCmd;
END_REGION

REGION Network 19: Transition for STATE Num:142 Tray Rdy to Drop Fix- Wait for Robot Accept request
   RUNG wire#powerrail
      Contact( #s142_TrayRdyDropFix )
      I_Contact( #sStWtResetRel )
      Contact( #sSst )
      Contact( #iR1DropOver )
      Coil( #s142_TrayRdyDropFix_T1 )
   END_RUNG
   // the same network as SCL:
   #s142_TrayRdyDropFix_T1 := #s142_TrayRdyDropFix AND NOT #sStWtResetRel AND #sSst AND #iR1DropOver;
END_REGION

REGION Network 20: STATE Num:142 Tray Rdy to Drop Fix- Wait for Robot Accept request
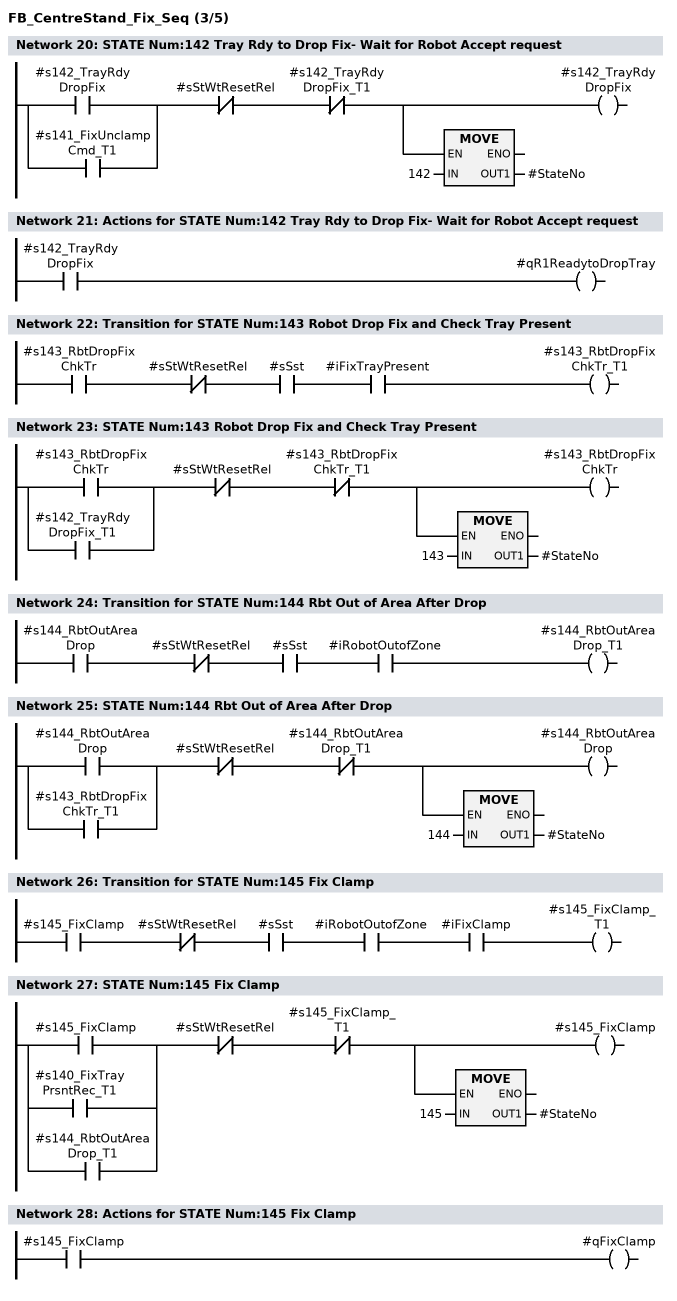
   RUNG wire#powerrail
      Contact( #s142_TrayRdyDropFix )
      wire#w1
      I_Contact( #sStWtResetRel )
      I_Contact( #s142_TrayRdyDropFix_T1 )
      wire#w2
      Coil( #s142_TrayRdyDropFix )
   END_RUNG
   RUNG wire#powerrail
      Contact( #s141_FixUnclampCmd_T1 )
   END_RUNG wire#w1
   RUNG wire#w2
      { S7_GenerateENO := "TRUE" } Move(in := 142, out1 => #StateNo)
   END_RUNG
   // the same network as SCL:
   #s142_TrayRdyDropFix := (#s142_TrayRdyDropFix OR #s141_FixUnclampCmd_T1) AND NOT #sStWtResetRel AND NOT #s142_TrayRdyDropFix_T1;
   IF #s142_TrayRdyDropFix THEN #StateNo := 142; END_IF;
END_REGION

REGION Network 21: Actions for STATE Num:142 Tray Rdy to Drop Fix- Wait for Robot Accept request
   RUNG wire#powerrail
      Contact( #s142_TrayRdyDropFix )
      Coil( #qR1ReadytoDropTray )
   END_RUNG
   // the same network as SCL:
   #qR1ReadytoDropTray := #s142_TrayRdyDropFix;
END_REGION

REGION Network 22: Transition for STATE Num:143 Robot Drop Fix and Check Tray Present
   RUNG wire#powerrail
      Contact( #s143_RbtDropFixChkTr )
      I_Contact( #sStWtResetRel )
      Contact( #sSst )
      Contact( #iFixTrayPresent )
      Coil( #s143_RbtDropFixChkTr_T1 )
   END_RUNG
   // the same network as SCL:
   #s143_RbtDropFixChkTr_T1 := #s143_RbtDropFixChkTr AND NOT #sStWtResetRel AND #sSst AND #iFixTrayPresent;
END_REGION

REGION Network 23: STATE Num:143 Robot Drop Fix and Check Tray Present
   RUNG wire#powerrail
      Contact( #s143_RbtDropFixChkTr )
      wire#w1
      I_Contact( #sStWtResetRel )
      I_Contact( #s143_RbtDropFixChkTr_T1 )
      wire#w2
      Coil( #s143_RbtDropFixChkTr )
   END_RUNG
   RUNG wire#powerrail
      Contact( #s142_TrayRdyDropFix_T1 )
   END_RUNG wire#w1
   RUNG wire#w2
      { S7_GenerateENO := "TRUE" } Move(in := 143, out1 => #StateNo)
   END_RUNG
   // the same network as SCL:
   #s143_RbtDropFixChkTr := (#s143_RbtDropFixChkTr OR #s142_TrayRdyDropFix_T1) AND NOT #sStWtResetRel AND NOT #s143_RbtDropFixChkTr_T1;
   IF #s143_RbtDropFixChkTr THEN #StateNo := 143; END_IF;
END_REGION

REGION Network 24: Transition for STATE Num:144 Rbt Out of Area After Drop
   RUNG wire#powerrail
      Contact( #s144_RbtOutAreaDrop )
      I_Contact( #sStWtResetRel )
      Contact( #sSst )
      Contact( #iRobotOutofZone )
      Coil( #s144_RbtOutAreaDrop_T1 )
   END_RUNG
   // the same network as SCL:
   #s144_RbtOutAreaDrop_T1 := #s144_RbtOutAreaDrop AND NOT #sStWtResetRel AND #sSst AND #iRobotOutofZone;
END_REGION

REGION Network 25: STATE Num:144 Rbt Out of Area After Drop
   RUNG wire#powerrail
      Contact( #s144_RbtOutAreaDrop )
      wire#w1
      I_Contact( #sStWtResetRel )
      I_Contact( #s144_RbtOutAreaDrop_T1 )
      wire#w2
      Coil( #s144_RbtOutAreaDrop )
   END_RUNG
   RUNG wire#powerrail
      Contact( #s143_RbtDropFixChkTr_T1 )
   END_RUNG wire#w1
   RUNG wire#w2
      { S7_GenerateENO := "TRUE" } Move(in := 144, out1 => #StateNo)
   END_RUNG
   // the same network as SCL:
   #s144_RbtOutAreaDrop := (#s144_RbtOutAreaDrop OR #s143_RbtDropFixChkTr_T1) AND NOT #sStWtResetRel AND NOT #s144_RbtOutAreaDrop_T1;
   IF #s144_RbtOutAreaDrop THEN #StateNo := 144; END_IF;
END_REGION

REGION Network 26: Transition for STATE Num:145 Fix Clamp
   RUNG wire#powerrail
      Contact( #s145_FixClamp )
      I_Contact( #sStWtResetRel )
      Contact( #sSst )
      Contact( #iRobotOutofZone )
      Contact( #iFixClamp )
      Coil( #s145_FixClamp_T1 )
   END_RUNG
   // the same network as SCL:
   #s145_FixClamp_T1 := #s145_FixClamp AND NOT #sStWtResetRel AND #sSst AND #iRobotOutofZone AND #iFixClamp;
END_REGION

REGION Network 27: STATE Num:145 Fix Clamp
   RUNG wire#powerrail
      Contact( #s145_FixClamp )
      wire#w1
      I_Contact( #sStWtResetRel )
      I_Contact( #s145_FixClamp_T1 )
      wire#w2
      Coil( #s145_FixClamp )
   END_RUNG
   RUNG wire#powerrail
      Contact( #s140_FixTrayPrsntRec_T1 )
   END_RUNG wire#w1
   RUNG wire#powerrail
      Contact( #s144_RbtOutAreaDrop_T1 )
   END_RUNG wire#w1
   RUNG wire#w2
      { S7_GenerateENO := "TRUE" } Move(in := 145, out1 => #StateNo)
   END_RUNG
   // the same network as SCL:
   #s145_FixClamp := (#s145_FixClamp OR #s140_FixTrayPrsntRec_T1 OR #s144_RbtOutAreaDrop_T1) AND NOT #sStWtResetRel AND NOT #s145_FixClamp_T1;
   IF #s145_FixClamp THEN #StateNo := 145; END_IF;
END_REGION

REGION Network 28: Actions for STATE Num:145 Fix Clamp
   RUNG wire#powerrail
      Contact( #s145_FixClamp )
      Coil( #qFixClamp )
   END_RUNG
   // the same network as SCL:
   #qFixClamp := #s145_FixClamp;
END_REGION

REGION Network 29: Transition for STATE Num:146 Robot-2 All Alloys Pick Or Drop Operation over
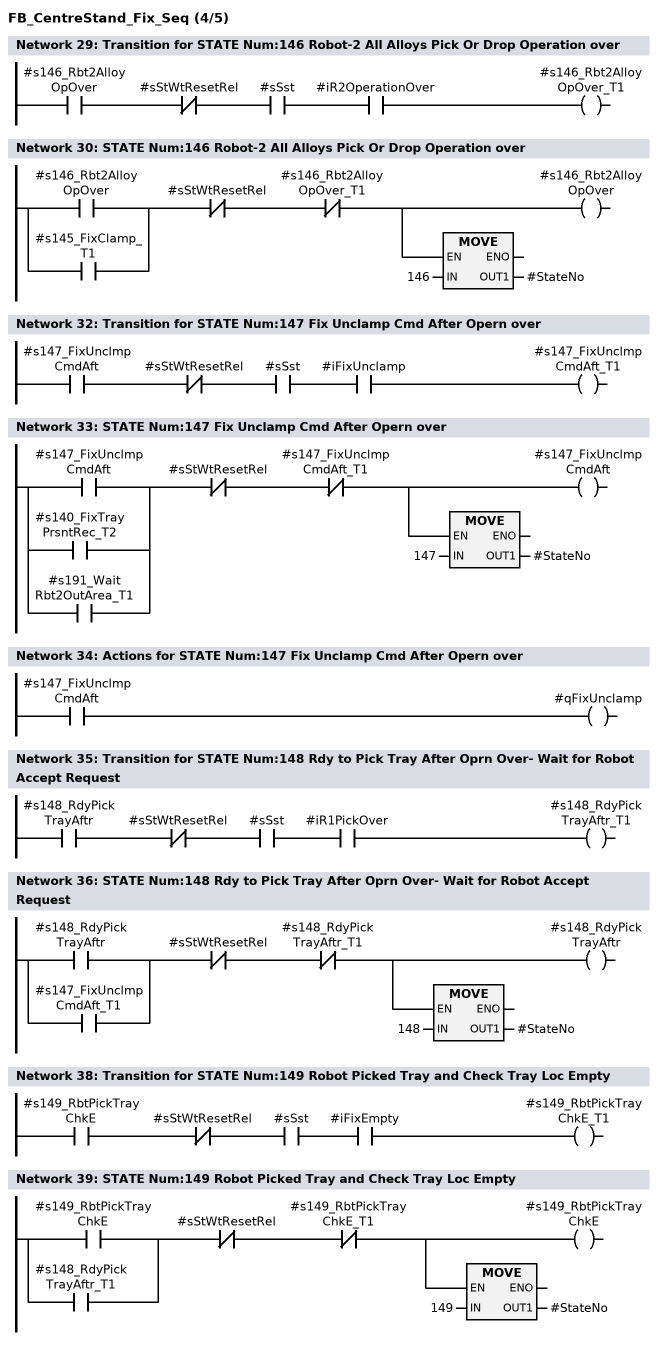
   RUNG wire#powerrail
      Contact( #s146_Rbt2AlloyOpOver )
      I_Contact( #sStWtResetRel )
      Contact( #sSst )
      Contact( #iR2OperationOver )
      Coil( #s146_Rbt2AlloyOpOver_T1 )
   END_RUNG
   // the same network as SCL:
   #s146_Rbt2AlloyOpOver_T1 := #s146_Rbt2AlloyOpOver AND NOT #sStWtResetRel AND #sSst AND #iR2OperationOver;
END_REGION

REGION Network 30: STATE Num:146 Robot-2 All Alloys Pick Or Drop Operation over
   RUNG wire#powerrail
      Contact( #s146_Rbt2AlloyOpOver )
      wire#w1
      I_Contact( #sStWtResetRel )
      I_Contact( #s146_Rbt2AlloyOpOver_T1 )
      wire#w2
      Coil( #s146_Rbt2AlloyOpOver )
   END_RUNG
   RUNG wire#powerrail
      Contact( #s145_FixClamp_T1 )
   END_RUNG wire#w1
   RUNG wire#w2
      { S7_GenerateENO := "TRUE" } Move(in := 146, out1 => #StateNo)
   END_RUNG
   // the same network as SCL:
   #s146_Rbt2AlloyOpOver := (#s146_Rbt2AlloyOpOver OR #s145_FixClamp_T1) AND NOT #sStWtResetRel AND NOT #s146_Rbt2AlloyOpOver_T1;
   IF #s146_Rbt2AlloyOpOver THEN #StateNo := 146; END_IF;
END_REGION

NETWORK
TITLE = Actions for STATE Num:146 Robot-2 All Alloys Pick Or Drop Operation over
      A     #s146_Rbt2AlloyOpOver;
      =     #qR2OperationStart;
      A     #s146_Rbt2AlloyOpOver;
      A     #iR2ServiceActivated;
      S     #iqR2ServiceActive;
      A     #s146_Rbt2AlloyOpOver;
      A     #iR2OperationOver;
      A     #iqR2ServiceActive;
      R     #iqR2ServiceActive;

REGION Network 32: Transition for STATE Num:147 Fix Unclamp Cmd After Opern over
   RUNG wire#powerrail
      Contact( #s147_FixUnclmpCmdAft )
      I_Contact( #sStWtResetRel )
      Contact( #sSst )
      Contact( #iFixUnclamp )
      Coil( #s147_FixUnclmpCmdAft_T1 )
   END_RUNG
   // the same network as SCL:
   #s147_FixUnclmpCmdAft_T1 := #s147_FixUnclmpCmdAft AND NOT #sStWtResetRel AND #sSst AND #iFixUnclamp;
END_REGION

REGION Network 33: STATE Num:147 Fix Unclamp Cmd After Opern over
   RUNG wire#powerrail
      Contact( #s147_FixUnclmpCmdAft )
      wire#w1
      I_Contact( #sStWtResetRel )
      I_Contact( #s147_FixUnclmpCmdAft_T1 )
      wire#w2
      Coil( #s147_FixUnclmpCmdAft )
   END_RUNG
   RUNG wire#powerrail
      Contact( #s140_FixTrayPrsntRec_T2 )
   END_RUNG wire#w1
   RUNG wire#powerrail
      Contact( #s191_WaitRbt2OutArea_T1 )
   END_RUNG wire#w1
   RUNG wire#w2
      { S7_GenerateENO := "TRUE" } Move(in := 147, out1 => #StateNo)
   END_RUNG
   // the same network as SCL:
   #s147_FixUnclmpCmdAft := (#s147_FixUnclmpCmdAft OR #s140_FixTrayPrsntRec_T2 OR #s191_WaitRbt2OutArea_T1) AND NOT #sStWtResetRel AND NOT #s147_FixUnclmpCmdAft_T1;
   IF #s147_FixUnclmpCmdAft THEN #StateNo := 147; END_IF;
END_REGION

REGION Network 34: Actions for STATE Num:147 Fix Unclamp Cmd After Opern over
   RUNG wire#powerrail
      Contact( #s147_FixUnclmpCmdAft )
      Coil( #qFixUnclamp )
   END_RUNG
   // the same network as SCL:
   #qFixUnclamp := #s147_FixUnclmpCmdAft;
END_REGION

REGION Network 35: Transition for STATE Num:148 Rdy to Pick Tray After Oprn Over- Wait for Robot Accept Request
   RUNG wire#powerrail
      Contact( #s148_RdyPickTrayAftr )
      I_Contact( #sStWtResetRel )
      Contact( #sSst )
      Contact( #iR1PickOver )
      Coil( #s148_RdyPickTrayAftr_T1 )
   END_RUNG
   // the same network as SCL:
   #s148_RdyPickTrayAftr_T1 := #s148_RdyPickTrayAftr AND NOT #sStWtResetRel AND #sSst AND #iR1PickOver;
END_REGION

REGION Network 36: STATE Num:148 Rdy to Pick Tray After Oprn Over- Wait for Robot Accept Request
   RUNG wire#powerrail
      Contact( #s148_RdyPickTrayAftr )
      wire#w1
      I_Contact( #sStWtResetRel )
      I_Contact( #s148_RdyPickTrayAftr_T1 )
      wire#w2
      Coil( #s148_RdyPickTrayAftr )
   END_RUNG
   RUNG wire#powerrail
      Contact( #s147_FixUnclmpCmdAft_T1 )
   END_RUNG wire#w1
   RUNG wire#w2
      { S7_GenerateENO := "TRUE" } Move(in := 148, out1 => #StateNo)
   END_RUNG
   // the same network as SCL:
   #s148_RdyPickTrayAftr := (#s148_RdyPickTrayAftr OR #s147_FixUnclmpCmdAft_T1) AND NOT #sStWtResetRel AND NOT #s148_RdyPickTrayAftr_T1;
   IF #s148_RdyPickTrayAftr THEN #StateNo := 148; END_IF;
END_REGION

NETWORK
TITLE = Actions for STATE Num:148 Rdy to Pick Tray After Oprn Over- Wait for Robot Accept Request
      A     #s148_RdyPickTrayAftr;
      =     #qR1ReadytoPickTray;
      A     #s148_RdyPickTrayAftr;
      A     #iR1PickOver;
      R     #iqR2ServiceCompleted;

REGION Network 38: Transition for STATE Num:149 Robot Picked Tray and Check Tray Loc Empty
   RUNG wire#powerrail
      Contact( #s149_RbtPickTrayChkE )
      I_Contact( #sStWtResetRel )
      Contact( #sSst )
      Contact( #iFixEmpty )
      Coil( #s149_RbtPickTrayChkE_T1 )
   END_RUNG
   // the same network as SCL:
   #s149_RbtPickTrayChkE_T1 := #s149_RbtPickTrayChkE AND NOT #sStWtResetRel AND #sSst AND #iFixEmpty;
END_REGION

REGION Network 39: STATE Num:149 Robot Picked Tray and Check Tray Loc Empty
   RUNG wire#powerrail
      Contact( #s149_RbtPickTrayChkE )
      wire#w1
      I_Contact( #sStWtResetRel )
      I_Contact( #s149_RbtPickTrayChkE_T1 )
      wire#w2
      Coil( #s149_RbtPickTrayChkE )
   END_RUNG
   RUNG wire#powerrail
      Contact( #s148_RdyPickTrayAftr_T1 )
   END_RUNG wire#w1
   RUNG wire#w2
      { S7_GenerateENO := "TRUE" } Move(in := 149, out1 => #StateNo)
   END_RUNG
   // the same network as SCL:
   #s149_RbtPickTrayChkE := (#s149_RbtPickTrayChkE OR #s148_RdyPickTrayAftr_T1) AND NOT #sStWtResetRel AND NOT #s149_RbtPickTrayChkE_T1;
   IF #s149_RbtPickTrayChkE THEN #StateNo := 149; END_IF;
END_REGION

REGION Network 40: Actions for STATE Num:149 Robot Picked Tray and Check Tray Loc Empty
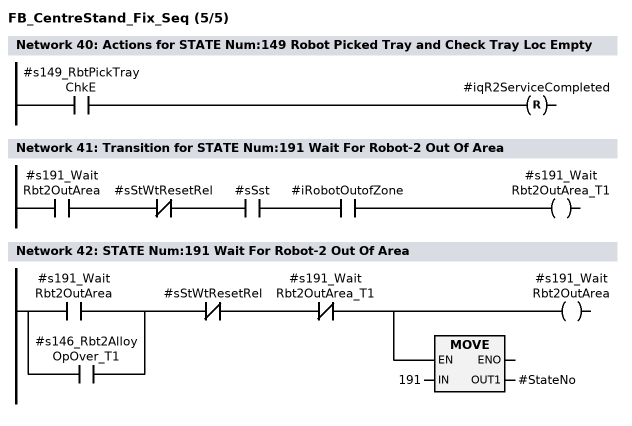
   RUNG wire#powerrail
      Contact( #s149_RbtPickTrayChkE )
      R_Coil( #iqR2ServiceCompleted )
   END_RUNG
   // the same network as SCL:
   IF #s149_RbtPickTrayChkE THEN #iqR2ServiceCompleted := FALSE; END_IF;
END_REGION

REGION Network 41: Transition for STATE Num:191 Wait For Robot-2 Out Of Area
   RUNG wire#powerrail
      Contact( #s191_WaitRbt2OutArea )
      I_Contact( #sStWtResetRel )
      Contact( #sSst )
      Contact( #iRobotOutofZone )
      Coil( #s191_WaitRbt2OutArea_T1 )
   END_RUNG
   // the same network as SCL:
   #s191_WaitRbt2OutArea_T1 := #s191_WaitRbt2OutArea AND NOT #sStWtResetRel AND #sSst AND #iRobotOutofZone;
END_REGION

REGION Network 42: STATE Num:191 Wait For Robot-2 Out Of Area
   RUNG wire#powerrail
      Contact( #s191_WaitRbt2OutArea )
      wire#w1
      I_Contact( #sStWtResetRel )
      I_Contact( #s191_WaitRbt2OutArea_T1 )
      wire#w2
      Coil( #s191_WaitRbt2OutArea )
   END_RUNG
   RUNG wire#powerrail
      Contact( #s146_Rbt2AlloyOpOver_T1 )
   END_RUNG wire#w1
   RUNG wire#w2
      { S7_GenerateENO := "TRUE" } Move(in := 191, out1 => #StateNo)
   END_RUNG
   // the same network as SCL:
   #s191_WaitRbt2OutArea := (#s191_WaitRbt2OutArea OR #s146_Rbt2AlloyOpOver_T1) AND NOT #sStWtResetRel AND NOT #s191_WaitRbt2OutArea_T1;
   IF #s191_WaitRbt2OutArea THEN #StateNo := 191; END_IF;
END_REGION
END_FUNCTION_BLOCK

FUNCTION_BLOCK "FB_GantryUnload_Seq"   // FB2, LAD
VERSION : 0.1
// stored: AutoNumber true, IsIECCheckEnabled false, UDAEnableTagReadback false
   VAR_INPUT
      iAutoRunning : Bool;
      iCenteringSlideAtHome : Bool;
      iCenteringSlideAtWork : Bool;
      iDistSenHighLimit : Int;
      iDistSenLowLimit : Int;
      iDistSensorIP : Int;
      iDryCycleWithoutPal : Bool;
      iGantryOutofZone : Bool;
      iGantryPickOver : Bool;
      iPCAckZero : Bool;
      iPCBypass : Bool;
      iPCDataReadOver : Bool;
      iPCDataWriteOver : Bool;
      iPalletPresent : Bool;
      iProcessStart : Bool;
      iReset_fault : Bool;
      iRetryPB : Bool;
      iScanErr : Bool;
      iScanOver : Bool;
      iScannerBypass : Bool;
      iSstMode : Bool;
      iSstPB : Bool;
   END_VAR
   VAR_OUTPUT
      qCenteringSlideAdvance : Bool;
      qCenteringSlideRetract : Bool;
      qCheckDistance : Bool;
      qGantryOkToUnload : Bool;
      qMsg : Array[0..2] of Bool;
      qPCReadCmd : Bool;
      qPCUploadCmd : Bool;
      qProcessOver : Bool;
      qScanCmd : Bool;
   END_VAR
   VAR DB_SPECIFIC
      StateNo : Int;
      s44_WaitResetRelease : Bool;
      s44_WaitResetRelease_T1 : Bool;
      s45_WaitGantryOutZone : Bool;
      s45_WaitGantryOutZone_T1 : Bool;
      s46_ChkStationHome : Bool;
      s46_ChkStationHome_T1 : Bool;
      s46_ChkStationHome_T2 : Bool;
      s47_WaitProcStartPZR : Bool;
      s47_WaitProcStartPZR_T1 : Bool;
      s48_ChkRecovery : Bool;
      s48_ChkRecovery_T1 : Bool;
      s48_ChkRecovery_T2 : Bool;
      s48_ChkRecovery_T3 : Bool;
      s49_WaitCentSlideAdv : Bool;
      s49_WaitCentSlideAdv_T1 : Bool;
      s50_WaitDistSensorFB : Bool;
      s50_WaitDistSensorFB_T1 : Bool;
      s51_WaitCentSlideRet : Bool;
      s51_WaitCentSlideRet_T1 : Bool;
      s52_WaitScanOver : Bool;
      s52_WaitScanOver_T1 : Bool;
      s52_WaitScanOver_T2 : Bool;
      s53_ChkDistOkWithPC : Bool;
      s53_ChkDistOkWithPC_T1 : Bool;
      s53_ChkDistOkWithPC_T2 : Bool;
      s54_WaitGantryUnload : Bool;
      s54_WaitGantryUnload_T1 : Bool;
      s55_WaitGantryUnldOvr : Bool;
      s55_WaitGantryUnldOvr_T1 : Bool;
      s56_WaitGantryOutZone : Bool;
      s56_WaitGantryOutZone_T1 : Bool;
      s57_ChkReelAbsentConv : Bool;
      s57_ChkReelAbsentConv_T1 : Bool;
      s58_WaitProcStartLow : Bool;
      s58_WaitProcStartLow_T1 : Bool;
      s61_ChkMeasDiamTol : Bool;
      s61_ChkMeasDiamTol_T1 : Bool;
      s61_ChkMeasDiamTol_T2 : Bool;
      s62_WaitPCAckZero : Bool;
      s62_WaitPCAckZero_T1 : Bool;
      s63_WaitDataWritePC : Bool;
      s63_WaitDataWritePC_T1 : Bool;
      s64_WaitOperatorIntv : Bool;
      s64_WaitOperatorIntv_T1 : Bool;
      s65_ChkScanRetryOver : Bool;
      s65_ChkScanRetryOver_T1 : Bool;
      s65_ChkScanRetryOver_T2 : Bool;
      s66_WaitOperatorDecis : Bool;
      s66_WaitOperatorDecis_T1 : Bool;
      s67_WaitCentSlideRet : Bool;
      s67_WaitCentSlideRet_T1 : Bool;
      s68_WaitPCAckZeroRead : Bool;
      s68_WaitPCAckZeroRead_T1 : Bool;
      s69_WaitDataReadPC : Bool;
      s69_WaitDataReadPC_T1 : Bool;
      sDistanceHighLimit : Int;
      sDistanceLowLimit : Int;
      sRecoveryInt : Int;
      sScanRetryCount : Int;
      sSst : Bool;
      sSstPulse : Bool;
      sSstRise : Bool;
   END_VAR
   VAR_TEMP
      tOne : Bool;
   END_VAR
   VAR_TEMP   // added for the SCL form of the ladder/FBD networks
      _w1 : Bool;
   END_VAR
BEGIN

REGION Network 1
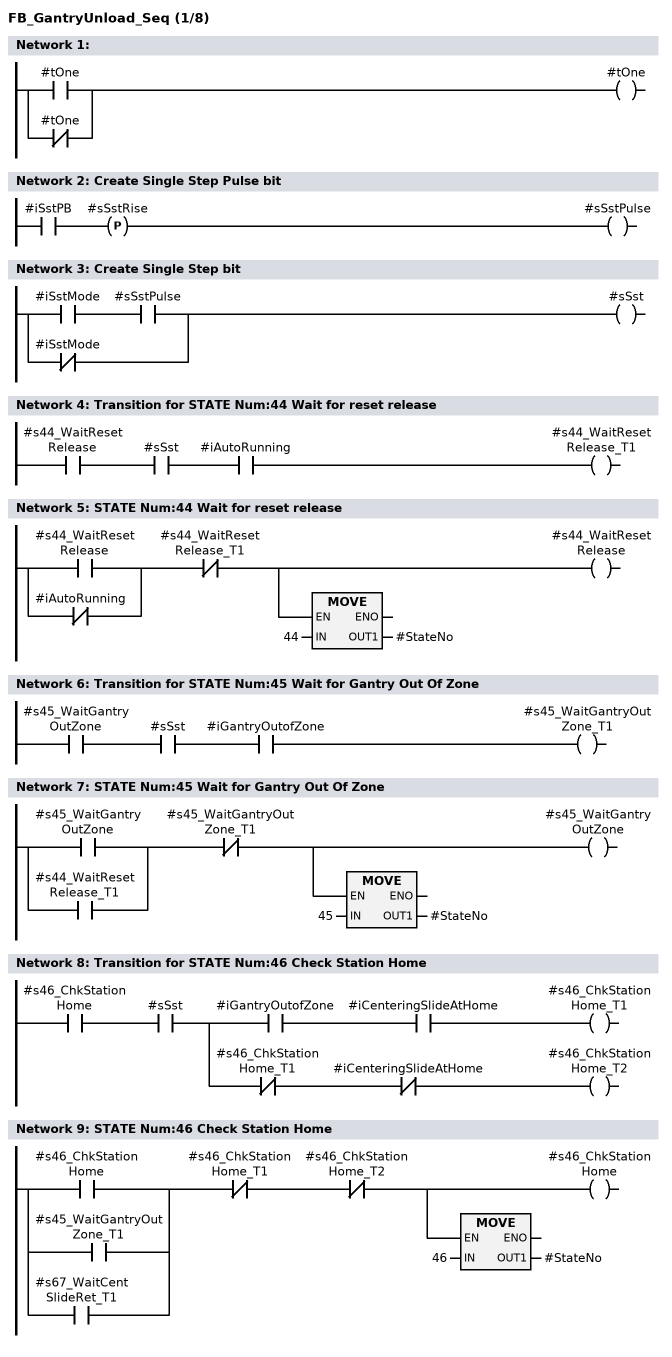
   RUNG wire#powerrail
      Contact( #tOne )
      wire#w1
      Coil( #tOne )
   END_RUNG
   RUNG wire#powerrail
      I_Contact( #tOne )
   END_RUNG wire#w1
   // the same network as SCL:
   #tOne := #tOne OR NOT #tOne;
END_REGION

REGION Network 2: Create Single Step Pulse bit
   RUNG wire#powerrail
      Contact( #iSstPB )
      P_Trig( #sSstRise )
      Coil( #sSstPulse )
   END_RUNG
   // the same network as SCL:
   #_w1 := #iSstPB AND NOT #sSstRise;   // rising edge
   #sSstRise := #iSstPB;
   #sSstPulse := #_w1;
END_REGION

REGION Network 3: Create Single Step bit
   RUNG wire#powerrail
      Contact( #iSstMode )
      Contact( #sSstPulse )
      wire#w1
      Coil( #sSst )
   END_RUNG
   RUNG wire#powerrail
      I_Contact( #iSstMode )
   END_RUNG wire#w1
   // the same network as SCL:
   #sSst := (#iSstMode AND #sSstPulse) OR NOT #iSstMode;
END_REGION

REGION Network 4: Transition for STATE Num:44 Wait for reset release
   RUNG wire#powerrail
      Contact( #s44_WaitResetRelease )
      Contact( #sSst )
      Contact( #iAutoRunning )
      Coil( #s44_WaitResetRelease_T1 )
   END_RUNG
   // the same network as SCL:
   #s44_WaitResetRelease_T1 := #s44_WaitResetRelease AND #sSst AND #iAutoRunning;
END_REGION

REGION Network 5: STATE Num:44 Wait for reset release
   RUNG wire#powerrail
      Contact( #s44_WaitResetRelease )
      wire#w1
      I_Contact( #s44_WaitResetRelease_T1 )
      wire#w2
      Coil( #s44_WaitResetRelease )
   END_RUNG
   RUNG wire#powerrail
      I_Contact( #iAutoRunning )
   END_RUNG wire#w1
   RUNG wire#w2
      { S7_GenerateENO := "TRUE" } Move(in := 44, out1 => #StateNo)
   END_RUNG
   // the same network as SCL:
   #s44_WaitResetRelease := (#s44_WaitResetRelease OR NOT #iAutoRunning) AND NOT #s44_WaitResetRelease_T1;
   IF #s44_WaitResetRelease THEN #StateNo := 44; END_IF;
END_REGION

REGION Network 6: Transition for STATE Num:45 Wait for Gantry Out Of Zone
   RUNG wire#powerrail
      Contact( #s45_WaitGantryOutZone )
      Contact( #sSst )
      Contact( #iGantryOutofZone )
      Coil( #s45_WaitGantryOutZone_T1 )
   END_RUNG
   // the same network as SCL:
   #s45_WaitGantryOutZone_T1 := #s45_WaitGantryOutZone AND #sSst AND #iGantryOutofZone;
END_REGION

REGION Network 7: STATE Num:45 Wait for Gantry Out Of Zone
   RUNG wire#powerrail
      Contact( #s45_WaitGantryOutZone )
      wire#w1
      I_Contact( #s45_WaitGantryOutZone_T1 )
      wire#w2
      Coil( #s45_WaitGantryOutZone )
   END_RUNG
   RUNG wire#powerrail
      Contact( #s44_WaitResetRelease_T1 )
   END_RUNG wire#w1
   RUNG wire#w2
      { S7_GenerateENO := "TRUE" } Move(in := 45, out1 => #StateNo)
   END_RUNG
   // the same network as SCL:
   #s45_WaitGantryOutZone := (#s45_WaitGantryOutZone OR #s44_WaitResetRelease_T1) AND NOT #s45_WaitGantryOutZone_T1;
   IF #s45_WaitGantryOutZone THEN #StateNo := 45; END_IF;
END_REGION

REGION Network 8: Transition for STATE Num:46 Check Station Home
   RUNG wire#powerrail
      Contact( #s46_ChkStationHome )
      Contact( #sSst )
      wire#w1
      Contact( #iGantryOutofZone )
      Contact( #iCenteringSlideAtHome )
      Coil( #s46_ChkStationHome_T1 )
   END_RUNG
   RUNG wire#w1
      I_Contact( #s46_ChkStationHome_T1 )
      I_Contact( #iCenteringSlideAtHome )
      Coil( #s46_ChkStationHome_T2 )
   END_RUNG
   // the same network as SCL:
   #_w1 := #s46_ChkStationHome AND #sSst;
   #s46_ChkStationHome_T1 := #_w1 AND #iGantryOutofZone AND #iCenteringSlideAtHome;
   #s46_ChkStationHome_T2 := #_w1 AND NOT #s46_ChkStationHome_T1 AND NOT #iCenteringSlideAtHome;
END_REGION

REGION Network 9: STATE Num:46 Check Station Home
   RUNG wire#powerrail
      Contact( #s46_ChkStationHome )
      wire#w1
      I_Contact( #s46_ChkStationHome_T1 )
      I_Contact( #s46_ChkStationHome_T2 )
      wire#w2
      Coil( #s46_ChkStationHome )
   END_RUNG
   RUNG wire#powerrail
      Contact( #s45_WaitGantryOutZone_T1 )
   END_RUNG wire#w1
   RUNG wire#powerrail
      Contact( #s67_WaitCentSlideRet_T1 )
   END_RUNG wire#w1
   RUNG wire#w2
      { S7_GenerateENO := "TRUE" } Move(in := 46, out1 => #StateNo)
   END_RUNG
   // the same network as SCL:
   #s46_ChkStationHome := (#s46_ChkStationHome OR #s45_WaitGantryOutZone_T1 OR #s67_WaitCentSlideRet_T1) AND NOT #s46_ChkStationHome_T1 AND NOT #s46_ChkStationHome_T2;
   IF #s46_ChkStationHome THEN #StateNo := 46; END_IF;
END_REGION

REGION Network 10: Transition for STATE Num:47 Wait for Process Start From PZR
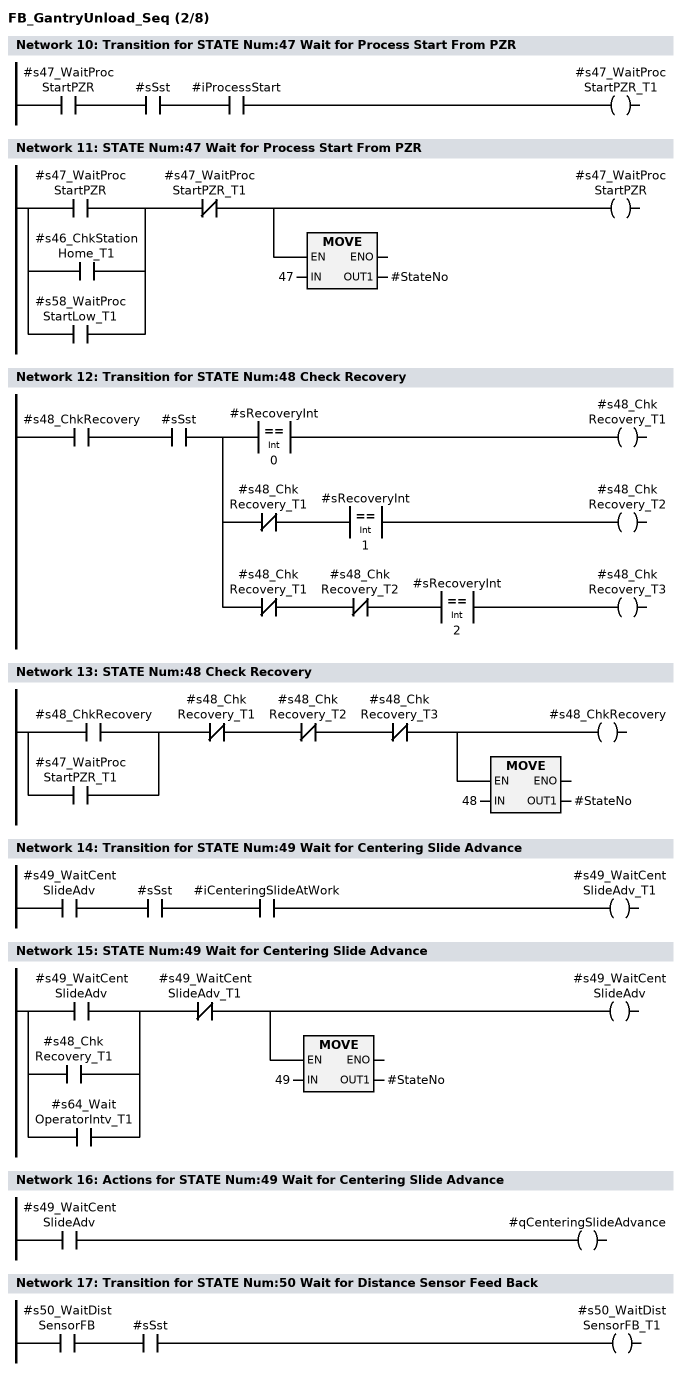
   RUNG wire#powerrail
      Contact( #s47_WaitProcStartPZR )
      Contact( #sSst )
      Contact( #iProcessStart )
      Coil( #s47_WaitProcStartPZR_T1 )
   END_RUNG
   // the same network as SCL:
   #s47_WaitProcStartPZR_T1 := #s47_WaitProcStartPZR AND #sSst AND #iProcessStart;
END_REGION

REGION Network 11: STATE Num:47 Wait for Process Start From PZR
   RUNG wire#powerrail
      Contact( #s47_WaitProcStartPZR )
      wire#w1
      I_Contact( #s47_WaitProcStartPZR_T1 )
      wire#w2
      Coil( #s47_WaitProcStartPZR )
   END_RUNG
   RUNG wire#powerrail
      Contact( #s46_ChkStationHome_T1 )
   END_RUNG wire#w1
   RUNG wire#powerrail
      Contact( #s58_WaitProcStartLow_T1 )
   END_RUNG wire#w1
   RUNG wire#w2
      { S7_GenerateENO := "TRUE" } Move(in := 47, out1 => #StateNo)
   END_RUNG
   // the same network as SCL:
   #s47_WaitProcStartPZR := (#s47_WaitProcStartPZR OR #s46_ChkStationHome_T1 OR #s58_WaitProcStartLow_T1) AND NOT #s47_WaitProcStartPZR_T1;
   IF #s47_WaitProcStartPZR THEN #StateNo := 47; END_IF;
END_REGION

REGION Network 12: Transition for STATE Num:48 Check Recovery
   RUNG wire#powerrail
      Contact( #s48_ChkRecovery )
      Contact( #sSst )
      wire#w1
      { S7_Templates := "SrcType := Int" } EQ_Contact(in1 := #sRecoveryInt, in2 := 0)
      Coil( #s48_ChkRecovery_T1 )
   END_RUNG
   RUNG wire#w1
      I_Contact( #s48_ChkRecovery_T1 )
      { S7_Templates := "SrcType := Int" } EQ_Contact(in1 := #sRecoveryInt, in2 := 1)
      Coil( #s48_ChkRecovery_T2 )
   END_RUNG
   RUNG wire#w1
      I_Contact( #s48_ChkRecovery_T1 )
      I_Contact( #s48_ChkRecovery_T2 )
      { S7_Templates := "SrcType := Int" } EQ_Contact(in1 := #sRecoveryInt, in2 := 2)
      Coil( #s48_ChkRecovery_T3 )
   END_RUNG
   // the same network as SCL:
   #_w1 := #s48_ChkRecovery AND #sSst;
   #s48_ChkRecovery_T1 := #_w1 AND (#sRecoveryInt = 0);
   #s48_ChkRecovery_T2 := #_w1 AND NOT #s48_ChkRecovery_T1 AND (#sRecoveryInt = 1);
   #s48_ChkRecovery_T3 := #_w1 AND NOT #s48_ChkRecovery_T1 AND NOT #s48_ChkRecovery_T2 AND (#sRecoveryInt = 2);
END_REGION

REGION Network 13: STATE Num:48 Check Recovery
   RUNG wire#powerrail
      Contact( #s48_ChkRecovery )
      wire#w1
      I_Contact( #s48_ChkRecovery_T1 )
      I_Contact( #s48_ChkRecovery_T2 )
      I_Contact( #s48_ChkRecovery_T3 )
      wire#w2
      Coil( #s48_ChkRecovery )
   END_RUNG
   RUNG wire#powerrail
      Contact( #s47_WaitProcStartPZR_T1 )
   END_RUNG wire#w1
   RUNG wire#w2
      { S7_GenerateENO := "TRUE" } Move(in := 48, out1 => #StateNo)
   END_RUNG
   // the same network as SCL:
   #s48_ChkRecovery := (#s48_ChkRecovery OR #s47_WaitProcStartPZR_T1) AND NOT #s48_ChkRecovery_T1 AND NOT #s48_ChkRecovery_T2 AND NOT #s48_ChkRecovery_T3;
   IF #s48_ChkRecovery THEN #StateNo := 48; END_IF;
END_REGION

REGION Network 14: Transition for STATE Num:49 Wait for Centering Slide Advance
   RUNG wire#powerrail
      Contact( #s49_WaitCentSlideAdv )
      Contact( #sSst )
      Contact( #iCenteringSlideAtWork )
      Coil( #s49_WaitCentSlideAdv_T1 )
   END_RUNG
   // the same network as SCL:
   #s49_WaitCentSlideAdv_T1 := #s49_WaitCentSlideAdv AND #sSst AND #iCenteringSlideAtWork;
END_REGION

REGION Network 15: STATE Num:49 Wait for Centering Slide Advance
   RUNG wire#powerrail
      Contact( #s49_WaitCentSlideAdv )
      wire#w1
      I_Contact( #s49_WaitCentSlideAdv_T1 )
      wire#w2
      Coil( #s49_WaitCentSlideAdv )
   END_RUNG
   RUNG wire#powerrail
      Contact( #s48_ChkRecovery_T1 )
   END_RUNG wire#w1
   RUNG wire#powerrail
      Contact( #s64_WaitOperatorIntv_T1 )
   END_RUNG wire#w1
   RUNG wire#w2
      { S7_GenerateENO := "TRUE" } Move(in := 49, out1 => #StateNo)
   END_RUNG
   // the same network as SCL:
   #s49_WaitCentSlideAdv := (#s49_WaitCentSlideAdv OR #s48_ChkRecovery_T1 OR #s64_WaitOperatorIntv_T1) AND NOT #s49_WaitCentSlideAdv_T1;
   IF #s49_WaitCentSlideAdv THEN #StateNo := 49; END_IF;
END_REGION

REGION Network 16: Actions for STATE Num:49 Wait for Centering Slide Advance
   RUNG wire#powerrail
      Contact( #s49_WaitCentSlideAdv )
      Coil( #qCenteringSlideAdvance )
   END_RUNG
   // the same network as SCL:
   #qCenteringSlideAdvance := #s49_WaitCentSlideAdv;
END_REGION

REGION Network 17: Transition for STATE Num:50 Wait for Distance Sensor Feed Back
   RUNG wire#powerrail
      Contact( #s50_WaitDistSensorFB )
      Contact( #sSst )
      Coil( #s50_WaitDistSensorFB_T1 )
   END_RUNG
   // the same network as SCL:
   #s50_WaitDistSensorFB_T1 := #s50_WaitDistSensorFB AND #sSst;
END_REGION

REGION Network 18: STATE Num:50 Wait for Distance Sensor Feed Back
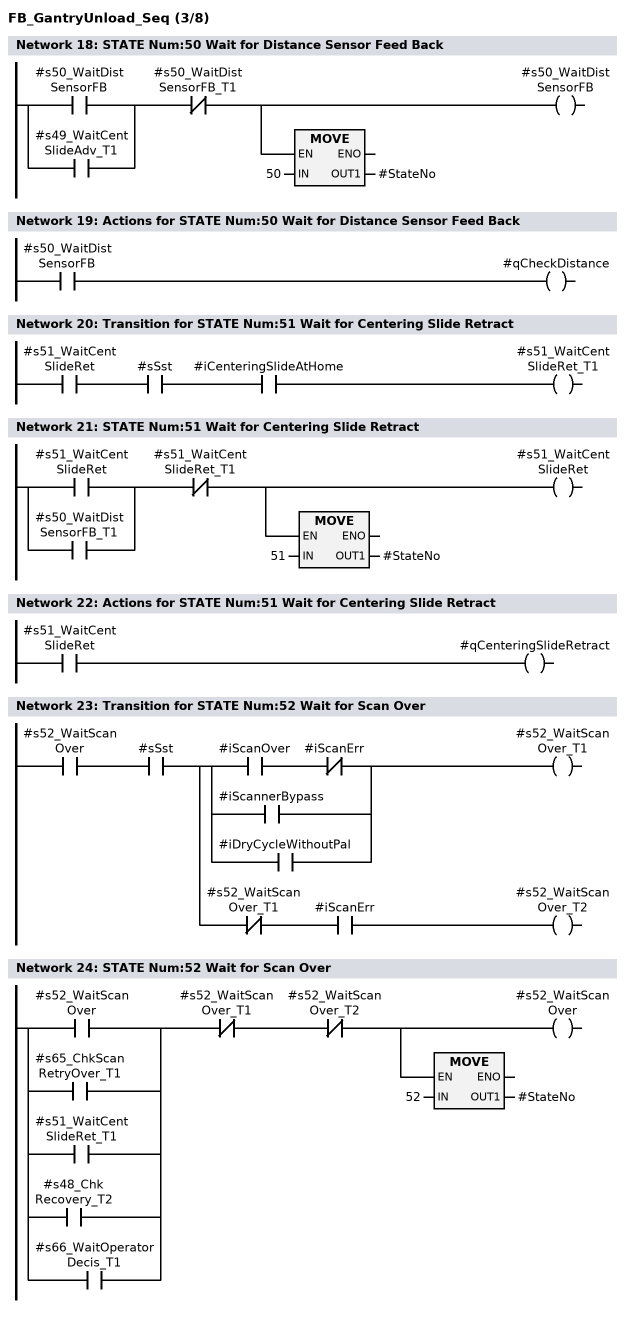
   RUNG wire#powerrail
      Contact( #s50_WaitDistSensorFB )
      wire#w1
      I_Contact( #s50_WaitDistSensorFB_T1 )
      wire#w2
      Coil( #s50_WaitDistSensorFB )
   END_RUNG
   RUNG wire#powerrail
      Contact( #s49_WaitCentSlideAdv_T1 )
   END_RUNG wire#w1
   RUNG wire#w2
      { S7_GenerateENO := "TRUE" } Move(in := 50, out1 => #StateNo)
   END_RUNG
   // the same network as SCL:
   #s50_WaitDistSensorFB := (#s50_WaitDistSensorFB OR #s49_WaitCentSlideAdv_T1) AND NOT #s50_WaitDistSensorFB_T1;
   IF #s50_WaitDistSensorFB THEN #StateNo := 50; END_IF;
END_REGION

REGION Network 19: Actions for STATE Num:50 Wait for Distance Sensor Feed Back
   RUNG wire#powerrail
      Contact( #s50_WaitDistSensorFB )
      Coil( #qCheckDistance )
   END_RUNG
   // the same network as SCL:
   #qCheckDistance := #s50_WaitDistSensorFB;
END_REGION

REGION Network 20: Transition for STATE Num:51 Wait for Centering Slide Retract
   RUNG wire#powerrail
      Contact( #s51_WaitCentSlideRet )
      Contact( #sSst )
      Contact( #iCenteringSlideAtHome )
      Coil( #s51_WaitCentSlideRet_T1 )
   END_RUNG
   // the same network as SCL:
   #s51_WaitCentSlideRet_T1 := #s51_WaitCentSlideRet AND #sSst AND #iCenteringSlideAtHome;
END_REGION

REGION Network 21: STATE Num:51 Wait for Centering Slide Retract
   RUNG wire#powerrail
      Contact( #s51_WaitCentSlideRet )
      wire#w1
      I_Contact( #s51_WaitCentSlideRet_T1 )
      wire#w2
      Coil( #s51_WaitCentSlideRet )
   END_RUNG
   RUNG wire#powerrail
      Contact( #s50_WaitDistSensorFB_T1 )
   END_RUNG wire#w1
   RUNG wire#w2
      { S7_GenerateENO := "TRUE" } Move(in := 51, out1 => #StateNo)
   END_RUNG
   // the same network as SCL:
   #s51_WaitCentSlideRet := (#s51_WaitCentSlideRet OR #s50_WaitDistSensorFB_T1) AND NOT #s51_WaitCentSlideRet_T1;
   IF #s51_WaitCentSlideRet THEN #StateNo := 51; END_IF;
END_REGION

REGION Network 22: Actions for STATE Num:51 Wait for Centering Slide Retract
   RUNG wire#powerrail
      Contact( #s51_WaitCentSlideRet )
      Coil( #qCenteringSlideRetract )
   END_RUNG
   // the same network as SCL:
   #qCenteringSlideRetract := #s51_WaitCentSlideRet;
END_REGION

REGION Network 23: Transition for STATE Num:52 Wait for Scan Over
   RUNG wire#powerrail
      Contact( #s52_WaitScanOver )
      Contact( #sSst )
      wire#w1
      Contact( #iScanOver )
      I_Contact( #iScanErr )
      wire#w2
      Coil( #s52_WaitScanOver_T1 )
   END_RUNG
   RUNG wire#w1
      Contact( #iScannerBypass )
   END_RUNG wire#w2
   RUNG wire#w1
      Contact( #iDryCycleWithoutPal )
   END_RUNG wire#w2
   RUNG wire#w1
      I_Contact( #s52_WaitScanOver_T1 )
      Contact( #iScanErr )
      Coil( #s52_WaitScanOver_T2 )
   END_RUNG
   // the same network as SCL:
   #_w1 := #s52_WaitScanOver AND #sSst;
   #s52_WaitScanOver_T1 := #_w1 AND ((#iScanOver AND NOT #iScanErr) OR #iScannerBypass OR #iDryCycleWithoutPal);
   #s52_WaitScanOver_T2 := #_w1 AND NOT #s52_WaitScanOver_T1 AND #iScanErr;
END_REGION

REGION Network 24: STATE Num:52 Wait for Scan Over
   RUNG wire#powerrail
      Contact( #s52_WaitScanOver )
      wire#w1
      I_Contact( #s52_WaitScanOver_T1 )
      I_Contact( #s52_WaitScanOver_T2 )
      wire#w2
      Coil( #s52_WaitScanOver )
   END_RUNG
   RUNG wire#powerrail
      Contact( #s65_ChkScanRetryOver_T1 )
   END_RUNG wire#w1
   RUNG wire#powerrail
      Contact( #s51_WaitCentSlideRet_T1 )
   END_RUNG wire#w1
   RUNG wire#powerrail
      Contact( #s48_ChkRecovery_T2 )
   END_RUNG wire#w1
   RUNG wire#powerrail
      Contact( #s66_WaitOperatorDecis_T1 )
   END_RUNG wire#w1
   RUNG wire#w2
      { S7_GenerateENO := "TRUE" } Move(in := 52, out1 => #StateNo)
   END_RUNG
   // the same network as SCL:
   #s52_WaitScanOver := (#s52_WaitScanOver OR #s65_ChkScanRetryOver_T1 OR #s51_WaitCentSlideRet_T1 OR #s48_ChkRecovery_T2 OR #s66_WaitOperatorDecis_T1) AND NOT #s52_WaitScanOver_T1 AND NOT #s52_WaitScanOver_T2;
   IF #s52_WaitScanOver THEN #StateNo := 52; END_IF;
END_REGION

REGION Network 25: Actions for STATE Num:52 Wait for Scan Over
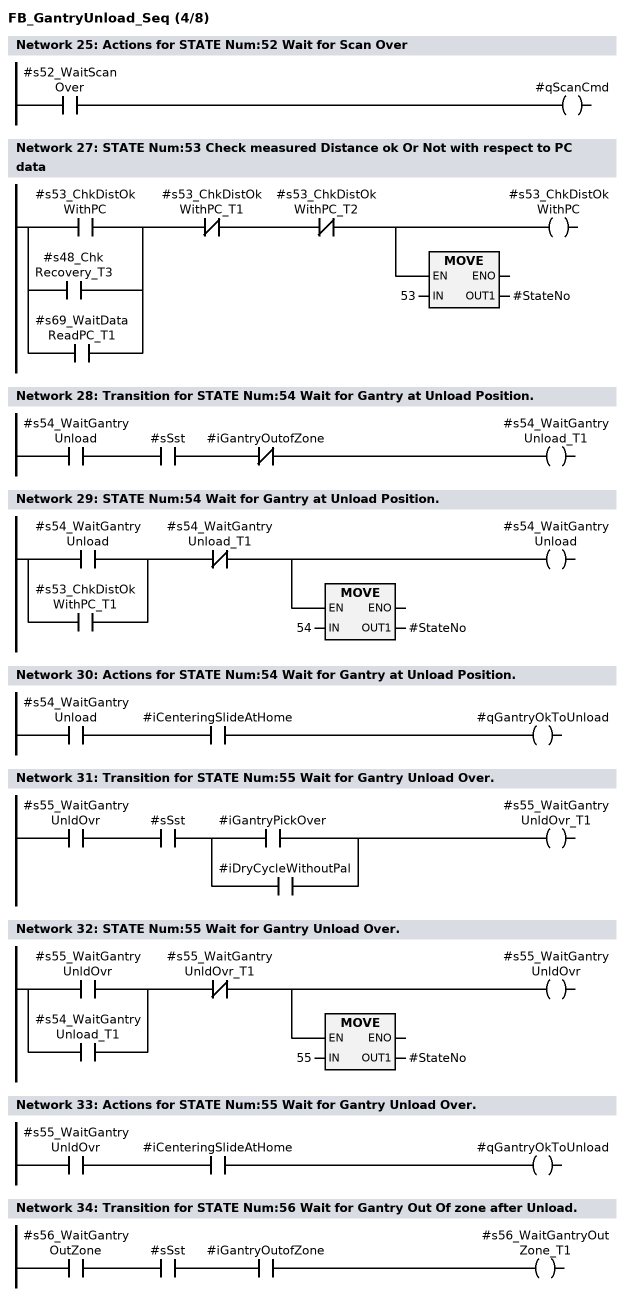
   RUNG wire#powerrail
      Contact( #s52_WaitScanOver )
      Coil( #qScanCmd )
   END_RUNG
   // the same network as SCL:
   #qScanCmd := #s52_WaitScanOver;
END_REGION

NETWORK
TITLE = Transition for STATE Num:53 Check measured Distance ok Or Not with respect to PC data
      A     #s53_ChkDistOkWithPC;
      A     #sSst;
      =     %L1.0;
      A     %L1.0;
      A(;
      L     #iDistSensorIP;
      L     #sDistanceLowLimit;
      >=R;
      );
      O(;
      L     #iDistSensorIP;
      L     #sDistanceHighLimit;
      <=R;
      );
      =     #s53_ChkDistOkWithPC_T1;
      A     %L1.0;
      AN    #s53_ChkDistOkWithPC_T1;
      A(;
      L     #iDistSensorIP;
      L     #sDistanceLowLimit;
      <R;
      );
      O(;
      L     #iDistSensorIP;
      L     #sDistanceHighLimit;
      >R;
      );
      =     #s53_ChkDistOkWithPC_T2;

REGION Network 27: STATE Num:53 Check measured Distance ok Or Not with respect to PC data
   RUNG wire#powerrail
      Contact( #s53_ChkDistOkWithPC )
      wire#w1
      I_Contact( #s53_ChkDistOkWithPC_T1 )
      I_Contact( #s53_ChkDistOkWithPC_T2 )
      wire#w2
      Coil( #s53_ChkDistOkWithPC )
   END_RUNG
   RUNG wire#powerrail
      Contact( #s48_ChkRecovery_T3 )
   END_RUNG wire#w1
   RUNG wire#powerrail
      Contact( #s69_WaitDataReadPC_T1 )
   END_RUNG wire#w1
   RUNG wire#w2
      { S7_GenerateENO := "TRUE" } Move(in := 53, out1 => #StateNo)
   END_RUNG
   // the same network as SCL:
   #s53_ChkDistOkWithPC := (#s53_ChkDistOkWithPC OR #s48_ChkRecovery_T3 OR #s69_WaitDataReadPC_T1) AND NOT #s53_ChkDistOkWithPC_T1 AND NOT #s53_ChkDistOkWithPC_T2;
   IF #s53_ChkDistOkWithPC THEN #StateNo := 53; END_IF;
END_REGION

REGION Network 28: Transition for STATE Num:54 Wait for Gantry at Unload Position.
   RUNG wire#powerrail
      Contact( #s54_WaitGantryUnload )
      Contact( #sSst )
      I_Contact( #iGantryOutofZone )
      Coil( #s54_WaitGantryUnload_T1 )
   END_RUNG
   // the same network as SCL:
   #s54_WaitGantryUnload_T1 := #s54_WaitGantryUnload AND #sSst AND NOT #iGantryOutofZone;
END_REGION

REGION Network 29: STATE Num:54 Wait for Gantry at Unload Position.
   RUNG wire#powerrail
      Contact( #s54_WaitGantryUnload )
      wire#w1
      I_Contact( #s54_WaitGantryUnload_T1 )
      wire#w2
      Coil( #s54_WaitGantryUnload )
   END_RUNG
   RUNG wire#powerrail
      Contact( #s53_ChkDistOkWithPC_T1 )
   END_RUNG wire#w1
   RUNG wire#w2
      { S7_GenerateENO := "TRUE" } Move(in := 54, out1 => #StateNo)
   END_RUNG
   // the same network as SCL:
   #s54_WaitGantryUnload := (#s54_WaitGantryUnload OR #s53_ChkDistOkWithPC_T1) AND NOT #s54_WaitGantryUnload_T1;
   IF #s54_WaitGantryUnload THEN #StateNo := 54; END_IF;
END_REGION

REGION Network 30: Actions for STATE Num:54 Wait for Gantry at Unload Position.
   RUNG wire#powerrail
      Contact( #s54_WaitGantryUnload )
      Contact( #iCenteringSlideAtHome )
      Coil( #qGantryOkToUnload )
   END_RUNG
   // the same network as SCL:
   #qGantryOkToUnload := #s54_WaitGantryUnload AND #iCenteringSlideAtHome;
END_REGION

REGION Network 31: Transition for STATE Num:55 Wait for Gantry Unload Over.
   RUNG wire#powerrail
      Contact( #s55_WaitGantryUnldOvr )
      Contact( #sSst )
      wire#w1
      Contact( #iGantryPickOver )
      wire#w2
      Coil( #s55_WaitGantryUnldOvr_T1 )
   END_RUNG
   RUNG wire#w1
      Contact( #iDryCycleWithoutPal )
   END_RUNG wire#w2
   // the same network as SCL:
   #s55_WaitGantryUnldOvr_T1 := #s55_WaitGantryUnldOvr AND #sSst AND (#iGantryPickOver OR #iDryCycleWithoutPal);
END_REGION

REGION Network 32: STATE Num:55 Wait for Gantry Unload Over.
   RUNG wire#powerrail
      Contact( #s55_WaitGantryUnldOvr )
      wire#w1
      I_Contact( #s55_WaitGantryUnldOvr_T1 )
      wire#w2
      Coil( #s55_WaitGantryUnldOvr )
   END_RUNG
   RUNG wire#powerrail
      Contact( #s54_WaitGantryUnload_T1 )
   END_RUNG wire#w1
   RUNG wire#w2
      { S7_GenerateENO := "TRUE" } Move(in := 55, out1 => #StateNo)
   END_RUNG
   // the same network as SCL:
   #s55_WaitGantryUnldOvr := (#s55_WaitGantryUnldOvr OR #s54_WaitGantryUnload_T1) AND NOT #s55_WaitGantryUnldOvr_T1;
   IF #s55_WaitGantryUnldOvr THEN #StateNo := 55; END_IF;
END_REGION

REGION Network 33: Actions for STATE Num:55 Wait for Gantry Unload Over.
   RUNG wire#powerrail
      Contact( #s55_WaitGantryUnldOvr )
      Contact( #iCenteringSlideAtHome )
      Coil( #qGantryOkToUnload )
   END_RUNG
   // the same network as SCL:
   #qGantryOkToUnload := #s55_WaitGantryUnldOvr AND #iCenteringSlideAtHome;
END_REGION

REGION Network 34: Transition for STATE Num:56 Wait for Gantry Out Of zone after Unload.
   RUNG wire#powerrail
      Contact( #s56_WaitGantryOutZone )
      Contact( #sSst )
      Contact( #iGantryOutofZone )
      Coil( #s56_WaitGantryOutZone_T1 )
   END_RUNG
   // the same network as SCL:
   #s56_WaitGantryOutZone_T1 := #s56_WaitGantryOutZone AND #sSst AND #iGantryOutofZone;
END_REGION

REGION Network 35: STATE Num:56 Wait for Gantry Out Of zone after Unload.
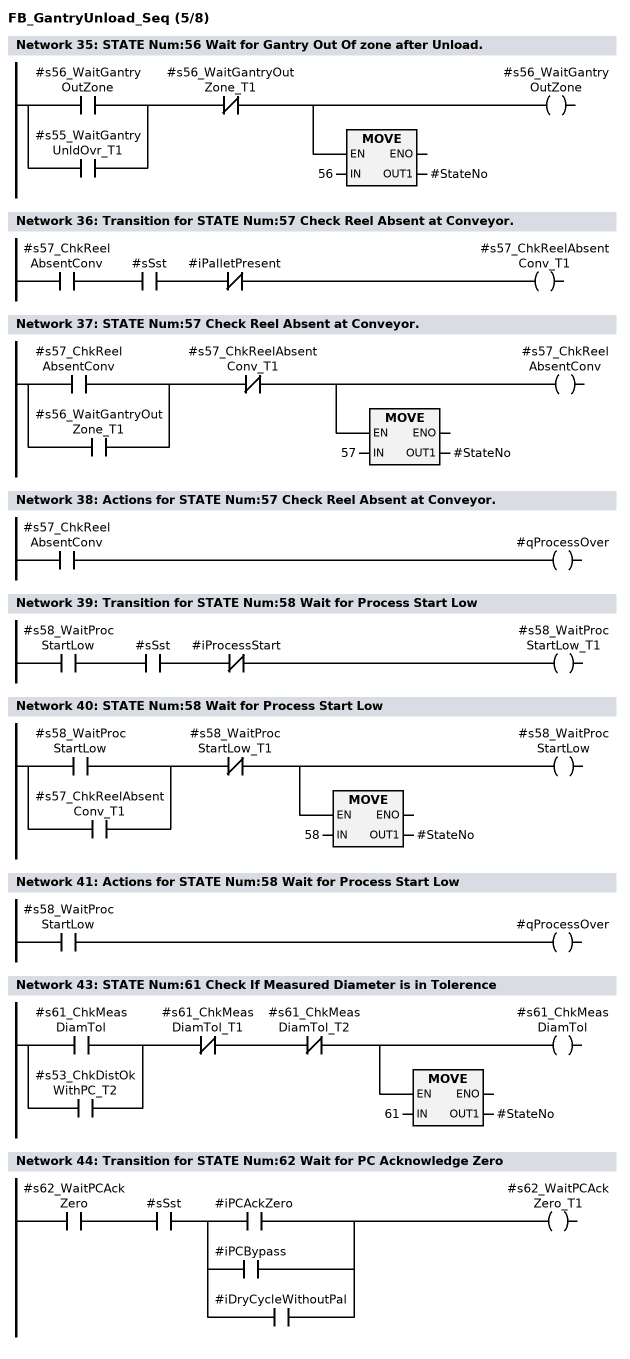
   RUNG wire#powerrail
      Contact( #s56_WaitGantryOutZone )
      wire#w1
      I_Contact( #s56_WaitGantryOutZone_T1 )
      wire#w2
      Coil( #s56_WaitGantryOutZone )
   END_RUNG
   RUNG wire#powerrail
      Contact( #s55_WaitGantryUnldOvr_T1 )
   END_RUNG wire#w1
   RUNG wire#w2
      { S7_GenerateENO := "TRUE" } Move(in := 56, out1 => #StateNo)
   END_RUNG
   // the same network as SCL:
   #s56_WaitGantryOutZone := (#s56_WaitGantryOutZone OR #s55_WaitGantryUnldOvr_T1) AND NOT #s56_WaitGantryOutZone_T1;
   IF #s56_WaitGantryOutZone THEN #StateNo := 56; END_IF;
END_REGION

REGION Network 36: Transition for STATE Num:57 Check Reel Absent at Conveyor.
   RUNG wire#powerrail
      Contact( #s57_ChkReelAbsentConv )
      Contact( #sSst )
      I_Contact( #iPalletPresent )
      Coil( #s57_ChkReelAbsentConv_T1 )
   END_RUNG
   // the same network as SCL:
   #s57_ChkReelAbsentConv_T1 := #s57_ChkReelAbsentConv AND #sSst AND NOT #iPalletPresent;
END_REGION

REGION Network 37: STATE Num:57 Check Reel Absent at Conveyor.
   RUNG wire#powerrail
      Contact( #s57_ChkReelAbsentConv )
      wire#w1
      I_Contact( #s57_ChkReelAbsentConv_T1 )
      wire#w2
      Coil( #s57_ChkReelAbsentConv )
   END_RUNG
   RUNG wire#powerrail
      Contact( #s56_WaitGantryOutZone_T1 )
   END_RUNG wire#w1
   RUNG wire#w2
      { S7_GenerateENO := "TRUE" } Move(in := 57, out1 => #StateNo)
   END_RUNG
   // the same network as SCL:
   #s57_ChkReelAbsentConv := (#s57_ChkReelAbsentConv OR #s56_WaitGantryOutZone_T1) AND NOT #s57_ChkReelAbsentConv_T1;
   IF #s57_ChkReelAbsentConv THEN #StateNo := 57; END_IF;
END_REGION

REGION Network 38: Actions for STATE Num:57 Check Reel Absent at Conveyor.
   RUNG wire#powerrail
      Contact( #s57_ChkReelAbsentConv )
      Coil( #qProcessOver )
   END_RUNG
   // the same network as SCL:
   #qProcessOver := #s57_ChkReelAbsentConv;
END_REGION

REGION Network 39: Transition for STATE Num:58 Wait for Process Start Low
   RUNG wire#powerrail
      Contact( #s58_WaitProcStartLow )
      Contact( #sSst )
      I_Contact( #iProcessStart )
      Coil( #s58_WaitProcStartLow_T1 )
   END_RUNG
   // the same network as SCL:
   #s58_WaitProcStartLow_T1 := #s58_WaitProcStartLow AND #sSst AND NOT #iProcessStart;
END_REGION

REGION Network 40: STATE Num:58 Wait for Process Start Low
   RUNG wire#powerrail
      Contact( #s58_WaitProcStartLow )
      wire#w1
      I_Contact( #s58_WaitProcStartLow_T1 )
      wire#w2
      Coil( #s58_WaitProcStartLow )
   END_RUNG
   RUNG wire#powerrail
      Contact( #s57_ChkReelAbsentConv_T1 )
   END_RUNG wire#w1
   RUNG wire#w2
      { S7_GenerateENO := "TRUE" } Move(in := 58, out1 => #StateNo)
   END_RUNG
   // the same network as SCL:
   #s58_WaitProcStartLow := (#s58_WaitProcStartLow OR #s57_ChkReelAbsentConv_T1) AND NOT #s58_WaitProcStartLow_T1;
   IF #s58_WaitProcStartLow THEN #StateNo := 58; END_IF;
END_REGION

REGION Network 41: Actions for STATE Num:58 Wait for Process Start Low
   RUNG wire#powerrail
      Contact( #s58_WaitProcStartLow )
      Coil( #qProcessOver )
   END_RUNG
   // the same network as SCL:
   #qProcessOver := #s58_WaitProcStartLow;
END_REGION

NETWORK
TITLE = Transition for STATE Num:61 Check If Measured Diameter is in Tolerence
      A     #s61_ChkMeasDiamTol;
      A     #sSst;
      =     %L1.0;
      A     %L1.0;
      A(;
      L     #iDistSenLowLimit;
      L     #iDistSensorIP;
      <=R;
      );
      O(;
      L     #iDistSensorIP;
      L     #iDistSenHighLimit;
      <=R;
      );
      =     #s61_ChkMeasDiamTol_T1;
      A     %L1.0;
      AN    #s61_ChkMeasDiamTol_T1;
      A(;
      L     #iDistSenLowLimit;
      L     #iDistSensorIP;
      >R;
      );
      O(;
      L     #iDistSensorIP;
      L     #iDistSenHighLimit;
      >R;
      );
      =     #s61_ChkMeasDiamTol_T2;

